// TIA Portal project "StdS71500PLCRack" (V17)

(* hardware
DEVICE "S7-1500/ET200MP-Station_1"  S7-1500 station
   slot 0: "Profilschiene_0"  Rack  6ES7 590-1***0-0AA0
   slot 1: "PLC_1"  CPU 1516-3 PN/DP  6ES7 516-3AN01-0AB0  V2.6
      slot 3: "CPU-Display_1"  6ES7591-1BA00-0AA0
      slot 32768: "PROFINET-Schnittstelle_1"  X1
      slot 33024: "PROFINET-Schnittstelle_2"  X2
      slot 33280: "DP-Schnittstelle_1"  X3
   slot 2: "DI 32x24VDC HF_1"  DI 32x24VDC HF  6ES7 521-1BL00-0AB0  V2.0
   slot 3: "DQ 32x24VDC/0.5A ST_1"  DQ 32x24VDC/0.5A ST  6ES7 522-1BL00-0AB0  V2.0
   slot 4: "AI 8xU/I/RTD/TC ST_1"  AI 8xU/I/RTD/TC ST  6ES7 531-7KF00-0AB0  V2.0
   slot 5: "AQ 4xU/I ST_1"  AQ 4xU/I ST  6ES7 532-5HD00-0AB0  V2.0
DEVICE "HMI_1"  TP700 Comfort
   slot 0: "HMI_1"  TP700 Comfort  6AV2 124-0GC01-0AX0  17.0.0.0
   slot 1: "HMI_RT_1"  TP700 Comfort  6AV2 124-0GC01-0AX0  17.0.0.0
   slot 5: "HMI_1.IE_CP_1"  PROFINET Interface  17.0.0.0
      slot 1: "PROFINET Interface_1"  PROFINET Interface
         slot 1: "Port_1"  Port
         slot 2: "Port_2"  Port
   slot 7: "HMI_1.MPI/DP_CP_1"  MPI/DP Interface  17.0.0.0
*)

// ===== PLC "PLC_1"  CPU 1516-3 PN/DP =====

VAR_GLOBAL   // PLC tag table "Standard-Variablentabelle"
   "System_Byte" AT %MB100 : Byte;
   "FirstScan" AT %M100.0 : Bool;
   "DiagStatusUpdate" AT %M100.1 : Bool;
   "AlwaysTRUE" AT %M100.2 : Bool;
   "AlwaysFALSE" AT %M100.3 : Bool;
   "Clock_Byte" AT %MB200 : Byte;
   "Clock_10Hz" AT %M200.0 : Bool;
   "Clock_5Hz" AT %M200.1 : Bool;
   "Clock_2.5Hz" AT %M200.2 : Bool;
   "Clock_2Hz" AT %M200.3 : Bool;
   "Clock_1.25Hz" AT %M200.4 : Bool;
   "Clock_1Hz" AT %M200.5 : Bool;
   "Clock_0.625Hz" AT %M200.6 : Bool;
   "Clock_0.5Hz" AT %M200.7 : Bool;
   "Tag_1" AT %M10.0 : Bool;
   "Tag_2" AT %M10.1 : Bool;
   "Tag_3" AT %M10.2 : Bool;
   "Tag_4" AT %M10.3 : Bool;
   "Tag_5" AT %M10.4 : Bool;
   "Tag_6" AT %M10.5 : Bool;
   "Tag_7" AT %M10.6 : Bool;
   "Tag_8" AT %M10.7 : Bool;
   "temp_AUTO_B" AT %M300.5 : Bool;
   "A_W_Testing" AT %M300.0 : Bool;
   "ACK_Status" AT %M300.2 : Bool;
   "Tag_11" AT %M300.3 : Bool;
   "Tag_9" AT %M300.7 : Bool;
   "Tag_10" AT %M11.0 : Bool;
   "Tag_12" AT %M11.1 : Bool;
   "Tag_13" AT %M11.2 : Bool;
END_VAR

DATA_BLOCK "PainMix_DB"   // DB1
{ S7_Optimized_Access := 'TRUE' }
VERSION : 0.1
   VAR
      Agitator_MainT : Int;
      Sol_1_Switch : Bool;
      Sol_1_Pipe1 : Int;
      Sol_1_Pipe2 : Int;
      RED_Pipe : Int;
      GREEN_Pipe : Int;
      BLUE_Pipe : Int;
      Control_Mode : Bool := false;
      Sol_1_ValveCont : Bool;
      Sol_1_Valve_Status : Bool;
      Sol_2_Valve_Status : Bool;
      Red_Valve_Status : Bool;
      Green_Valve_Status : Bool;
      Blue_Valve_Status : Bool;
      MainTank_Mixer_Status : Bool;
      Sol_2_ValveCont : Bool;
      Red_ValveCont : Bool;
      Green_ValveCont : Bool;
      Blue_ValveCont : Bool;
      Red_P_Rotor : Int;
      Green_P_Rotor : Int;
      Blue_P_Rotor : Int;
      Red_Tank_Level : Int := 40;
      Blue_Tank_Level : Int := 40;
      Green_Tank_Level : Int := 40;
      Sol_1_Tank_Level : Int := 40;
      Sol_2_Tank_Level : Int := 40;
      MainTank_Mixer_Cont : Bool;
      MainTank_Tank_Level : Int := 40;
      AUTO_Mode : Bool;
      AUTO_Mode_Prior : Int;
      temp_Auto_1 : Bool;
      Alarm_ACK : Bool;
   END_VAR
BEGIN
END_DATA_BLOCK

DATA_BLOCK "Paramters_Paint_Mix"   // DB7
{ S7_Optimized_Access := 'TRUE' }
VERSION : 0.1
   VAR
      ResinE_Flow_Act : Real := 1.6;
      ResinE_Flow_Set : Real := 1.8;
      Defoaming_Set : Real := 3.6;
      "Gloss Ratio_Set" : Real := 34.5;
      Binder_Flow_Act : Real := 2.2;
      Binder_Flow_Set : Real := 2.5;
      Level_Set_R : Real := 13.5;
      Level_Set_G : Real := 13.5;
      Level_Set_B : Real := 13.5;
      Flowrate_Set_R : Real := 3.1;
      Flowrate_Set_G : Real := 3.1;
      Flowrate_Set_B : Real := 3.1;
      Viscosity_Set_R : Real := 2.1;
      Viscosity_Set_G : Real := 2.7;
      Viscosity_Set_B : Real := 3.1;
      Density_Set_R : Real := 1.4;
      Density_Set_G : Real := 1.5;
      Density_Set_B : Real := 1.7;
      Temperature_Set_R : Real := 88.5;
      Temperature_Set_G : Real := 88.5;
      Temperature_Set_B : Real := 88.5;
      Pressure_Set_R : Real := 6.6;
      Pressure_Set_G : Real := 6.6;
      Pressure_Set_B : Real := 6.6;
      MixingSpeed_Set_MT : Real := 33.5;
      pH_MT : Real := 8.7;
      Viscosity_Set_MT : Real := 2.9;
      Level_Set_MT : Real := 17.0;
      Act_Red_Tank_Temp : Real := 73.5;
      Act_Green_Tank_Temp : Real := 76.2;
      Act_Blue_Tank_Temp : Real := 77.5;
      Act_Red_Tank_Press : Real := 5.3;
      Act_Green_Tank_Press : Real := 6.1;
      Act_Blue_Tank_Press : Real := 5.9;
      Recipe_Name : String := 'Pearl Gray';
      Recipe_ID : String := '001';
      Equip_ID : String := 'TN15112';
      Batch_ID : String := '052B';
      Batch_Size : String := '85 litr';
      Start_Time : String := '28/01/2025, 14:56:32';
      Alarm_1 : Bool;
      Alarm_2 : Bool;
      Warning_1 : Bool;
      Warning_2 : Bool;
      Warning_3 : Bool;
      "Common_A-W" : Bool;
      Language : Bool := false;
      Button_Language : Bool;
      MainOverview : Bool;
      Parameters : Bool;
      RecipeM : Bool;
      UserM : Bool;
      AlarmSt : Bool;
      IOSt : Bool;
   END_VAR
BEGIN
END_DATA_BLOCK

DATA_BLOCK "DI"   // DB8
{ S7_Optimized_Access := 'TRUE' }
VERSION : 0.1
   VAR
      "I0.0" : Bool;
      "I0.1" : Bool := true;
      "I0.2" : Bool;
      "I0.3" : Bool := true;
      "I0.4" : Bool;
      "I0.5" : Bool;
      "I0.6" : Bool := true;
      "I0.7" : Bool;
      "I1.0" : Bool;
      "I1.1" : Bool;
      "I1.2" : Bool;
      "I1.3" : Bool := true;
      "I1.4" : Bool;
      "I1.5" : Bool;
      "I1.6" : Bool;
      "I1.7" : Bool := true;
      "I2.0" : Bool := true;
      "I2.1" : Bool;
      "I2.2" : Bool;
      "I2.3" : Bool := true;
   END_VAR
BEGIN
END_DATA_BLOCK

DATA_BLOCK "DO"   // DB9
{ S7_Optimized_Access := 'TRUE' }
VERSION : 0.1
   VAR
      "Q0.0" : Bool;
      "Q0.1" : Bool;
      "Q0.2" : Bool;
      "Q0.3" : Bool;
      "Q0.4" : Bool;
      "Q0.5" : Bool;
      "Q0.6" : Bool;
      "Q0.7" : Bool;
      "Q1.0" : Bool;
      "Q1.1" : Bool;
      "Q1.2" : Bool;
      "Q1.3" : Bool;
      "Q1.4" : Bool;
      "Q1.5" : Bool;
      "Q1.6" : Bool;
      "Q1.7" : Bool := true;
      "Q2.0" : Bool;
      "Q2.1" : Bool;
      "Q2.2" : Bool := true;
      "Q2.3" : Bool := true;
   END_VAR
BEGIN
END_DATA_BLOCK

DATA_BLOCK "Recipe"   // DB10
{ S7_Optimized_Access := 'TRUE' }
VERSION : 0.1
   VAR
      "Pigment Concentration" : Real;
      "Resin Type and Ratio" : Real;
      "Solvent Composition" : Real;
      "Additive Ratios" : Real;
      "Drying Agent Ratio" : Real;
      "Viscosity Target" : Real;
      "Gloss Level" : Real;
      "pH Control Range" : Real;
      "Mixing Time" : Real;
      "Curing Agent Proportion" : Real;
      Recipe_Name : String;
   END_VAR
BEGIN
END_DATA_BLOCK

// folder: System blocks/Program resources

DATA_BLOCK "IEC_Timer_0_DB"   // DB2
{ S7_Optimized_Access := 'TRUE' }
AUTHOR : Simatic
FAMILY : IEC
NAME : IEC_TMR
VERSION : 1.0
// stored: InstanceOfName IEC_TIMER
"IEC_TIMER"
BEGIN
END_DATA_BLOCK

DATA_BLOCK "IEC_Timer_0_DB_1"   // DB3
{ S7_Optimized_Access := 'TRUE' }
AUTHOR : Simatic
FAMILY : IEC
NAME : IEC_TMR
VERSION : 1.0
// stored: InstanceOfName IEC_TIMER
"IEC_TIMER"
BEGIN
END_DATA_BLOCK

DATA_BLOCK "IEC_Timer_0_DB_2"   // DB4
{ S7_Optimized_Access := 'TRUE' }
AUTHOR : Simatic
FAMILY : IEC
NAME : IEC_TMR
VERSION : 1.0
// stored: InstanceOfName IEC_TIMER
"IEC_TIMER"
BEGIN
END_DATA_BLOCK

DATA_BLOCK "IEC_Timer_0_DB_3"   // DB5
{ S7_Optimized_Access := 'TRUE' }
AUTHOR : Simatic
FAMILY : IEC
NAME : IEC_TMR
VERSION : 1.0
// stored: InstanceOfName IEC_TIMER
"IEC_TIMER"
BEGIN
END_DATA_BLOCK

DATA_BLOCK "IEC_Timer_0_DB_4"   // DB6
{ S7_Optimized_Access := 'TRUE' }
AUTHOR : Simatic
FAMILY : IEC
NAME : IEC_TMR
VERSION : 1.0
// stored: InstanceOfName IEC_TIMER
"IEC_TIMER"
BEGIN
END_DATA_BLOCK

DATA_BLOCK "IEC_Timer_0_DB_5"   // DB11
{ S7_Optimized_Access := 'TRUE' }
AUTHOR : Simatic
FAMILY : IEC
NAME : IEC_TMR
VERSION : 1.0
// stored: InstanceOfName IEC_TIMER
"IEC_TIMER"
BEGIN
END_DATA_BLOCK

DATA_BLOCK "IEC_Counter_0_DB"   // DB12
{ S7_Optimized_Access := 'TRUE' }
AUTHOR : Simatic
FAMILY : IEC
NAME : CNTR
VERSION : 1.0
// stored: InstanceOfName IEC_COUNTER
"IEC_COUNTER"
BEGIN
END_DATA_BLOCK

DATA_BLOCK "IEC_Timer_0_DB_6"   // DB13
{ S7_Optimized_Access := 'TRUE' }
AUTHOR : Simatic
FAMILY : IEC
NAME : IEC_TMR
VERSION : 1.0
// stored: InstanceOfName IEC_TIMER
"IEC_TIMER"
BEGIN
END_DATA_BLOCK

// folder: (top level)

ORGANIZATION_BLOCK "Main"   // OB1, LAD, ProgramCycle
TITLE = "Main Program Sweep (Cycle)"
{ S7_Optimized_Access := 'TRUE' }
VERSION : 0.1
   VAR_INPUT
      Initial_Call : Bool;   // Initial call of this OB
      Remanence : Bool;   // =True, if remanent data are available
   END_VAR
   VAR_TEMP   // added for the SCL form of the ladder/FBD networks
      _w1 : Bool;
      _w2 : Bool;
   END_VAR
BEGIN

REGION Network 1: AUTO Sequence Logic
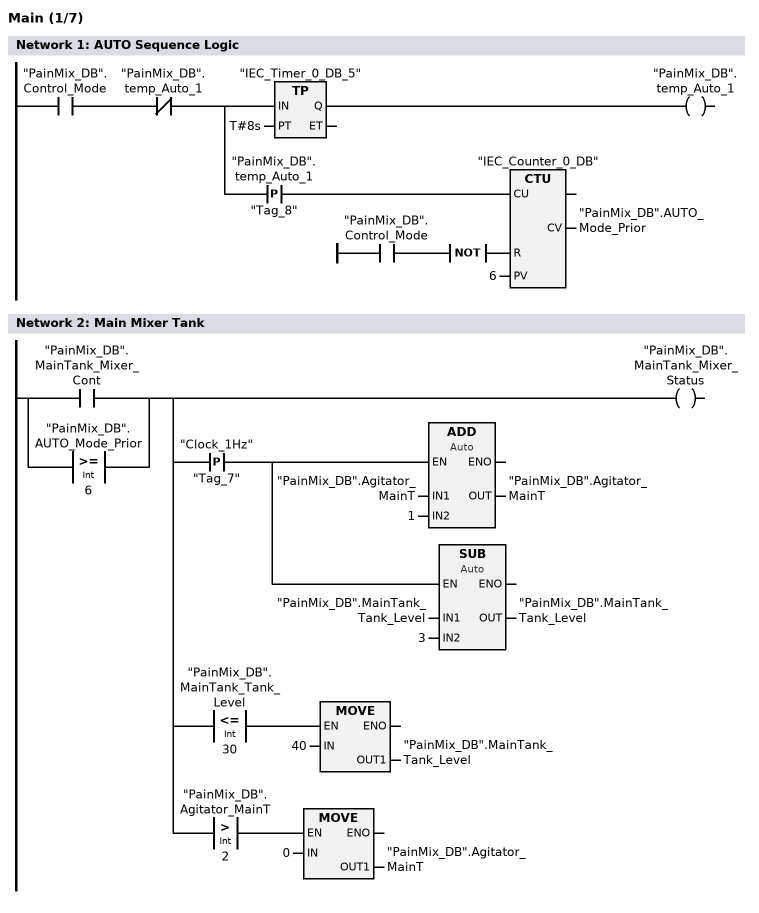
   #_w1 := "PainMix_DB".Control_Mode AND NOT "PainMix_DB".temp_Auto_1;
   "IEC_Timer_0_DB_5".TP(IN := #_w1, PT := T#8s);
   "PainMix_DB".temp_Auto_1 := "IEC_Timer_0_DB_5".Q;
   #_w2 := #_w1 AND "PainMix_DB".temp_Auto_1 AND NOT "Tag_8";   // rising edge of "PainMix_DB".temp_Auto_1
   "Tag_8" := "PainMix_DB".temp_Auto_1;
   "IEC_Counter_0_DB".CTU(CU := #_w2,
                          R := NOT "PainMix_DB".Control_Mode,
                          PV := 6,
                          CV => "PainMix_DB".AUTO_Mode_Prior);
END_REGION

REGION Network 2: Main Mixer Tank
   RUNG wire#powerrail
      Contact( "PainMix_DB".MainTank_Mixer_Cont )
      wire#w1
      Coil( "PainMix_DB".MainTank_Mixer_Status )
   END_RUNG
   RUNG wire#powerrail
      { S7_Templates := "SrcType := Int" } GE_Contact(in1 := "PainMix_DB".AUTO_Mode_Prior, in2 := 6)
   END_RUNG wire#w1
   RUNG wire#w1
      P_Contact(operand := "Clock_1Hz", bit := "Tag_7")
      wire#w2
      Add(in1 := "PainMix_DB".Agitator_MainT, in2 := 1, out => "PainMix_DB".Agitator_MainT)
   END_RUNG
   RUNG wire#w2
      Sub(in1 := "PainMix_DB".MainTank_Tank_Level, in2 := 3, out => "PainMix_DB".MainTank_Tank_Level)
   END_RUNG
   RUNG wire#w1
      { S7_Templates := "SrcType := Int" } LE_Contact(in1 := "PainMix_DB".MainTank_Tank_Level, in2 := 30)
      Move(in := 40, out1 => "PainMix_DB".MainTank_Tank_Level)
   END_RUNG
   RUNG wire#w1
      { S7_Templates := "SrcType := Int" } GT_Contact(in1 := "PainMix_DB".Agitator_MainT, in2 := 2)
      Move(in := 0, out1 => "PainMix_DB".Agitator_MainT)
   END_RUNG
   // the same network as SCL:
   "PainMix_DB".MainTank_Mixer_Status := "PainMix_DB".MainTank_Mixer_Cont OR ("PainMix_DB".AUTO_Mode_Prior >= 6);
   #_w1 := "PainMix_DB".MainTank_Mixer_Status AND "Clock_1Hz" AND NOT "Tag_7";   // rising edge of "Clock_1Hz"
   "Tag_7" := "Clock_1Hz";
   IF #_w1 THEN
       "PainMix_DB".Agitator_MainT := "PainMix_DB".Agitator_MainT + 1;
       "PainMix_DB".MainTank_Tank_Level := "PainMix_DB".MainTank_Tank_Level - 3;
   END_IF;
   IF "PainMix_DB".MainTank_Mixer_Status AND ("PainMix_DB".MainTank_Tank_Level <= 30) THEN
       "PainMix_DB".MainTank_Tank_Level := 40;
   END_IF;
   IF "PainMix_DB".MainTank_Mixer_Status AND ("PainMix_DB".Agitator_MainT > 2) THEN
       "PainMix_DB".Agitator_MainT := 0;
   END_IF;
END_REGION

REGION Network 3: Resin Solution
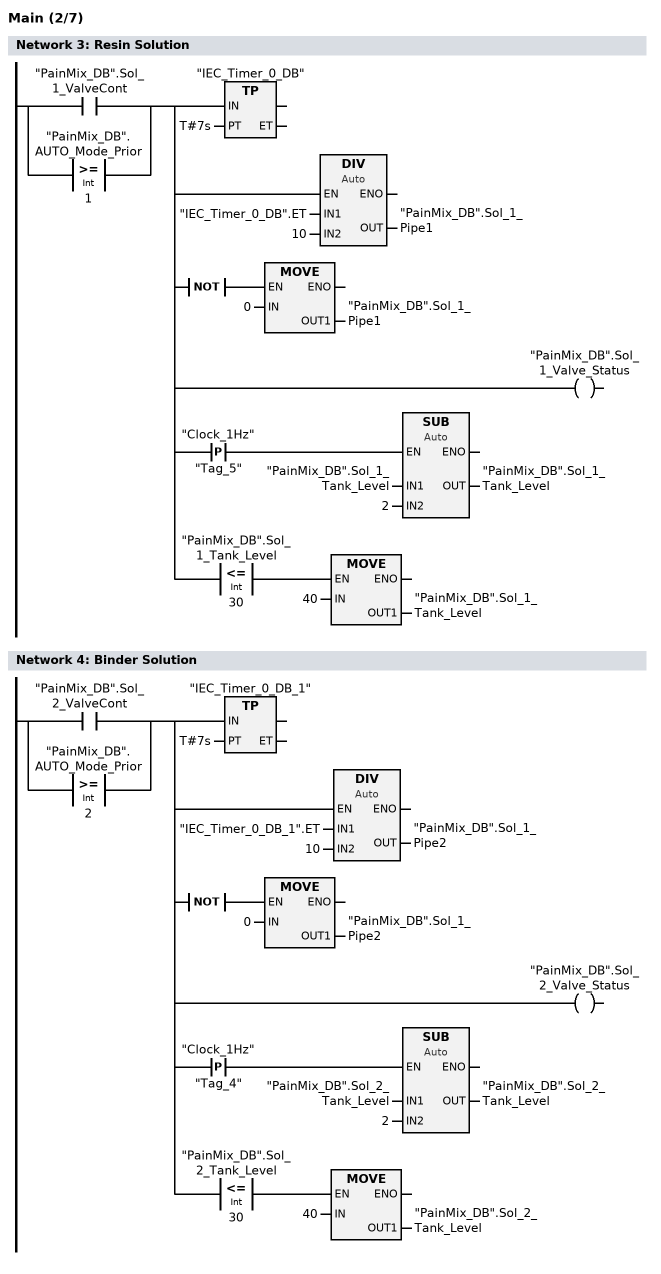
   #_w1 := "PainMix_DB".Sol_1_ValveCont OR ("PainMix_DB".AUTO_Mode_Prior >= 1);
   "IEC_Timer_0_DB".TP(IN := #_w1, PT := T#7s);
   IF #_w1 THEN "PainMix_DB".Sol_1_Pipe1 := "IEC_Timer_0_DB".ET / 10; END_IF;
   IF NOT #_w1 THEN "PainMix_DB".Sol_1_Pipe1 := 0; END_IF;
   "PainMix_DB".Sol_1_Valve_Status := #_w1;
   #_w2 := #_w1 AND "Clock_1Hz" AND NOT "Tag_5";   // rising edge of "Clock_1Hz"
   "Tag_5" := "Clock_1Hz";
   IF #_w2 THEN "PainMix_DB".Sol_1_Tank_Level := "PainMix_DB".Sol_1_Tank_Level - 2; END_IF;
   IF #_w1 AND ("PainMix_DB".Sol_1_Tank_Level <= 30) THEN "PainMix_DB".Sol_1_Tank_Level := 40; END_IF;
END_REGION

REGION Network 4: Binder Solution
   #_w1 := "PainMix_DB".Sol_2_ValveCont OR ("PainMix_DB".AUTO_Mode_Prior >= 2);
   "IEC_Timer_0_DB_1".TP(IN := #_w1, PT := T#7s);
   IF #_w1 THEN "PainMix_DB".Sol_1_Pipe2 := "IEC_Timer_0_DB_1".ET / 10; END_IF;
   IF NOT #_w1 THEN "PainMix_DB".Sol_1_Pipe2 := 0; END_IF;
   "PainMix_DB".Sol_2_Valve_Status := #_w1;
   #_w2 := #_w1 AND "Clock_1Hz" AND NOT "Tag_4";   // rising edge of "Clock_1Hz"
   "Tag_4" := "Clock_1Hz";
   IF #_w2 THEN "PainMix_DB".Sol_2_Tank_Level := "PainMix_DB".Sol_2_Tank_Level - 2; END_IF;
   IF #_w1 AND ("PainMix_DB".Sol_2_Tank_Level <= 30) THEN "PainMix_DB".Sol_2_Tank_Level := 40; END_IF;
END_REGION

REGION Network 5: RED
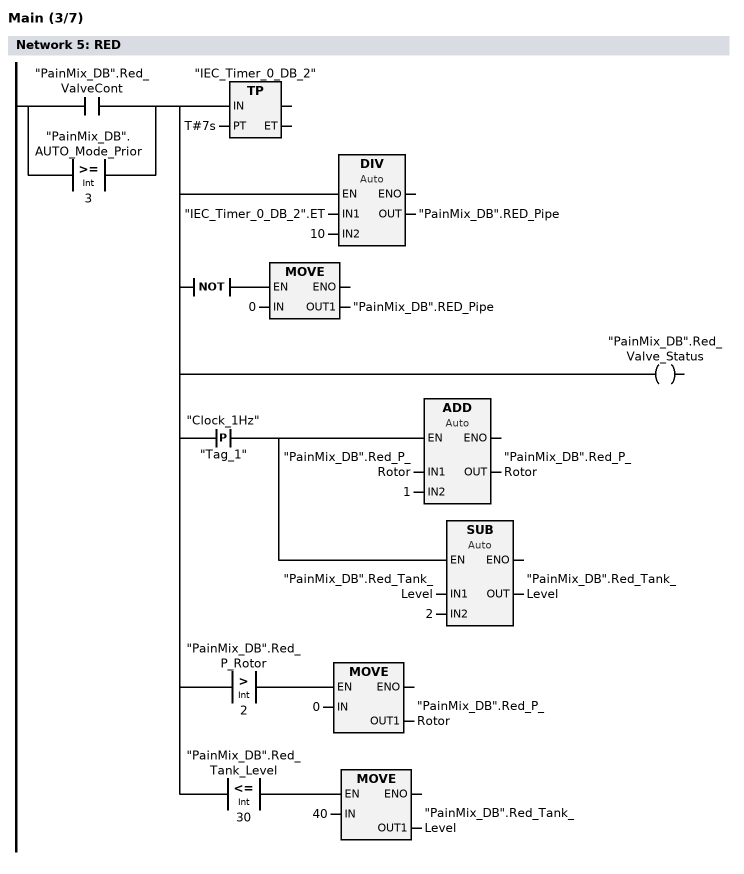
   #_w1 := "PainMix_DB".Red_ValveCont OR ("PainMix_DB".AUTO_Mode_Prior >= 3);
   "IEC_Timer_0_DB_2".TP(IN := #_w1, PT := T#7s);
   IF #_w1 THEN "PainMix_DB".RED_Pipe := "IEC_Timer_0_DB_2".ET / 10; END_IF;
   IF NOT #_w1 THEN "PainMix_DB".RED_Pipe := 0; END_IF;
   "PainMix_DB".Red_Valve_Status := #_w1;
   #_w2 := #_w1 AND "Clock_1Hz" AND NOT "Tag_1";   // rising edge of "Clock_1Hz"
   "Tag_1" := "Clock_1Hz";
   IF #_w2 THEN
       "PainMix_DB".Red_P_Rotor := "PainMix_DB".Red_P_Rotor + 1;
       "PainMix_DB".Red_Tank_Level := "PainMix_DB".Red_Tank_Level - 2;
   END_IF;
   IF #_w1 AND ("PainMix_DB".Red_P_Rotor > 2) THEN "PainMix_DB".Red_P_Rotor := 0; END_IF;
   IF #_w1 AND ("PainMix_DB".Red_Tank_Level <= 30) THEN "PainMix_DB".Red_Tank_Level := 40; END_IF;
END_REGION

REGION Network 6: GREEN
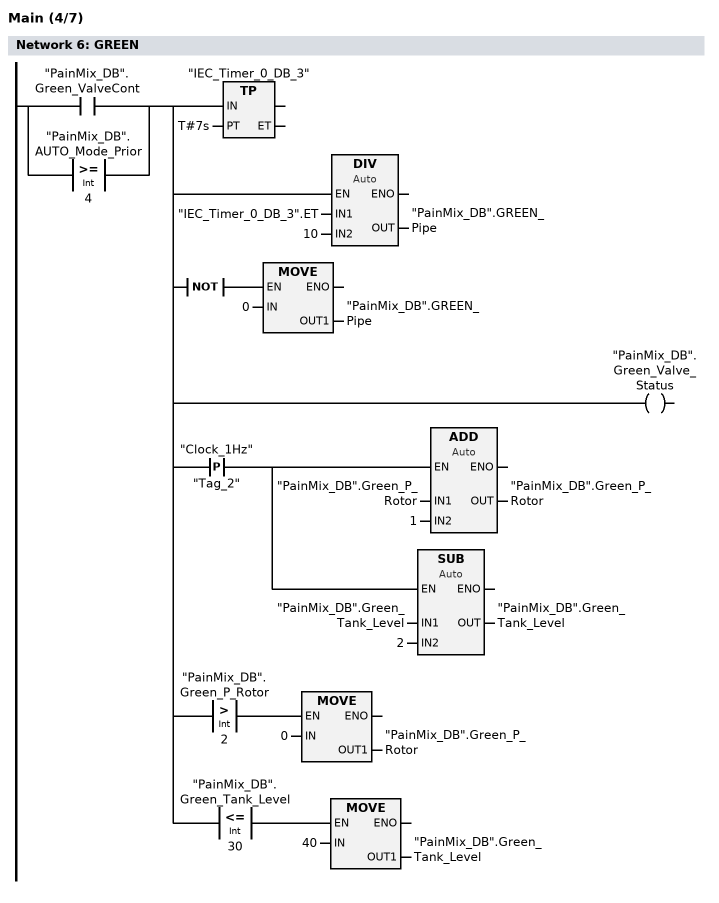
   #_w1 := "PainMix_DB".Green_ValveCont OR ("PainMix_DB".AUTO_Mode_Prior >= 4);
   "IEC_Timer_0_DB_3".TP(IN := #_w1, PT := T#7s);
   IF #_w1 THEN "PainMix_DB".GREEN_Pipe := "IEC_Timer_0_DB_3".ET / 10; END_IF;
   IF NOT #_w1 THEN "PainMix_DB".GREEN_Pipe := 0; END_IF;
   "PainMix_DB".Green_Valve_Status := #_w1;
   #_w2 := #_w1 AND "Clock_1Hz" AND NOT "Tag_2";   // rising edge of "Clock_1Hz"
   "Tag_2" := "Clock_1Hz";
   IF #_w2 THEN
       "PainMix_DB".Green_P_Rotor := "PainMix_DB".Green_P_Rotor + 1;
       "PainMix_DB".Green_Tank_Level := "PainMix_DB".Green_Tank_Level - 2;
   END_IF;
   IF #_w1 AND ("PainMix_DB".Green_P_Rotor > 2) THEN "PainMix_DB".Green_P_Rotor := 0; END_IF;
   IF #_w1 AND ("PainMix_DB".Green_Tank_Level <= 30) THEN "PainMix_DB".Green_Tank_Level := 40; END_IF;
END_REGION

REGION Network 7: BLUE
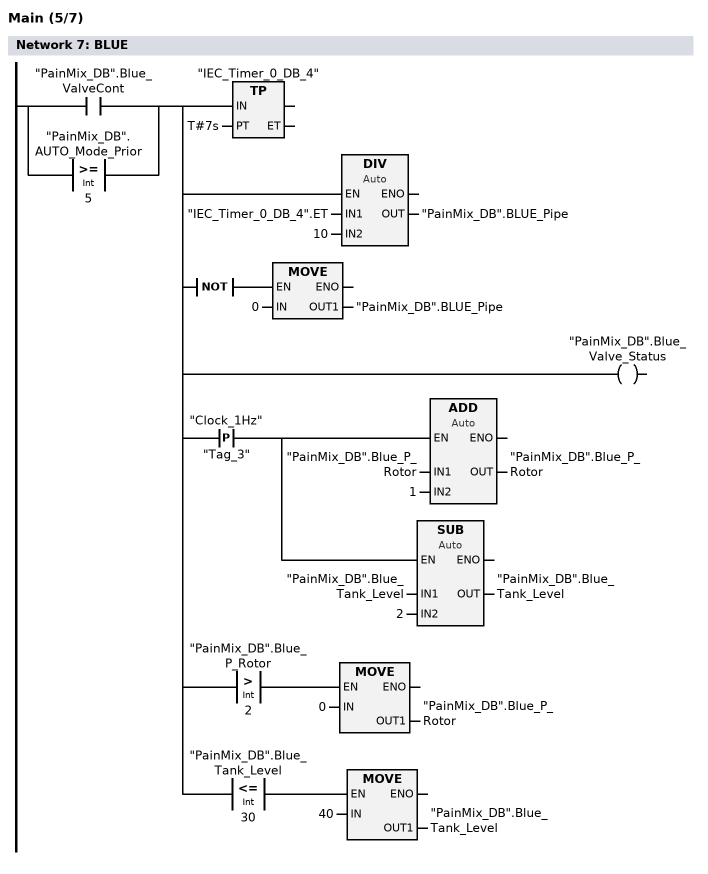
   #_w1 := "PainMix_DB".Blue_ValveCont OR ("PainMix_DB".AUTO_Mode_Prior >= 5);
   "IEC_Timer_0_DB_4".TP(IN := #_w1, PT := T#7s);
   IF #_w1 THEN "PainMix_DB".BLUE_Pipe := "IEC_Timer_0_DB_4".ET / 10; END_IF;
   IF NOT #_w1 THEN "PainMix_DB".BLUE_Pipe := 0; END_IF;
   "PainMix_DB".Blue_Valve_Status := #_w1;
   #_w2 := #_w1 AND "Clock_1Hz" AND NOT "Tag_3";   // rising edge of "Clock_1Hz"
   "Tag_3" := "Clock_1Hz";
   IF #_w2 THEN
       "PainMix_DB".Blue_P_Rotor := "PainMix_DB".Blue_P_Rotor + 1;
       "PainMix_DB".Blue_Tank_Level := "PainMix_DB".Blue_Tank_Level - 2;
   END_IF;
   IF #_w1 AND ("PainMix_DB".Blue_P_Rotor > 2) THEN "PainMix_DB".Blue_P_Rotor := 0; END_IF;
   IF #_w1 AND ("PainMix_DB".Blue_Tank_Level <= 30) THEN "PainMix_DB".Blue_Tank_Level := 40; END_IF;
END_REGION

REGION Network 8: Flucuation of Temp & Press of Tanks
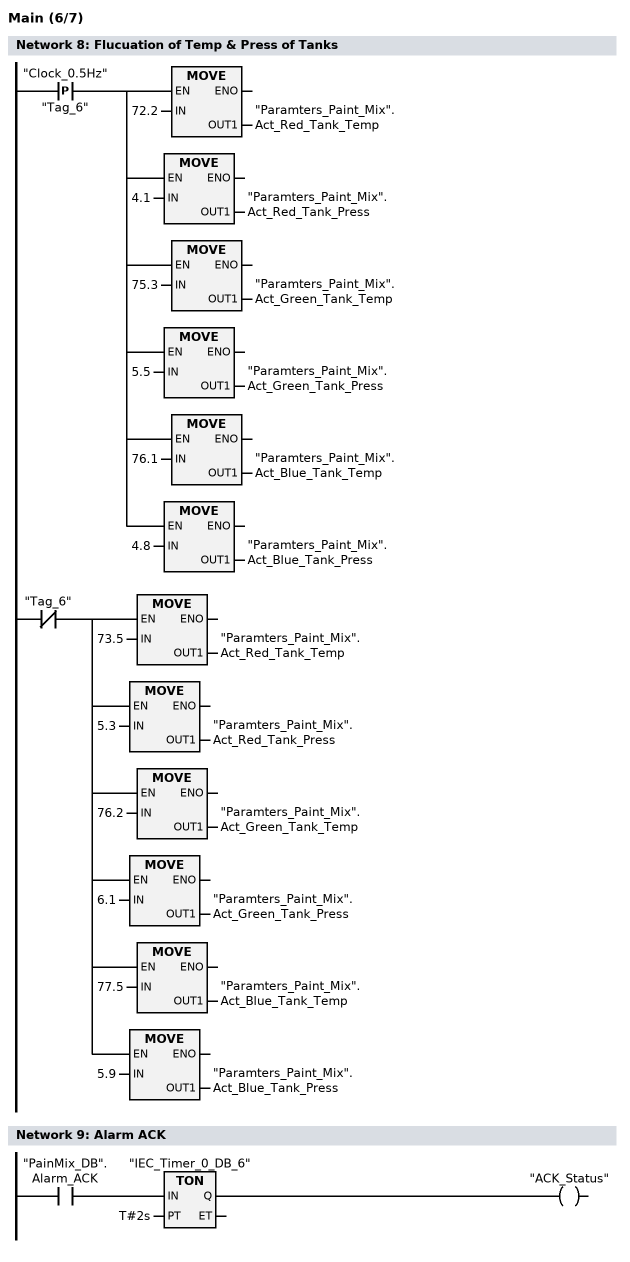
   RUNG wire#powerrail
      P_Contact(operand := "Clock_0.5Hz", bit := "Tag_6")
      wire#w1
      Move(in := 72.2, out1 => "Paramters_Paint_Mix".Act_Red_Tank_Temp)
   END_RUNG
   RUNG wire#w1
      Move(in := 4.1, out1 => "Paramters_Paint_Mix".Act_Red_Tank_Press)
   END_RUNG
   RUNG wire#w1
      Move(in := 75.3, out1 => "Paramters_Paint_Mix".Act_Green_Tank_Temp)
   END_RUNG
   RUNG wire#w1
      Move(in := 5.5, out1 => "Paramters_Paint_Mix".Act_Green_Tank_Press)
   END_RUNG
   RUNG wire#w1
      Move(in := 76.1, out1 => "Paramters_Paint_Mix".Act_Blue_Tank_Temp)
   END_RUNG
   RUNG wire#w1
      Move(in := 4.8, out1 => "Paramters_Paint_Mix".Act_Blue_Tank_Press)
   END_RUNG
   RUNG wire#powerrail
      I_Contact( "Tag_6" )
      wire#w2
      Move(in := 73.5, out1 => "Paramters_Paint_Mix".Act_Red_Tank_Temp)
   END_RUNG
   RUNG wire#w2
      Move(in := 5.3, out1 => "Paramters_Paint_Mix".Act_Red_Tank_Press)
   END_RUNG
   RUNG wire#w2
      Move(in := 76.2, out1 => "Paramters_Paint_Mix".Act_Green_Tank_Temp)
   END_RUNG
   RUNG wire#w2
      Move(in := 6.1, out1 => "Paramters_Paint_Mix".Act_Green_Tank_Press)
   END_RUNG
   RUNG wire#w2
      Move(in := 77.5, out1 => "Paramters_Paint_Mix".Act_Blue_Tank_Temp)
   END_RUNG
   RUNG wire#w2
      Move(in := 5.9, out1 => "Paramters_Paint_Mix".Act_Blue_Tank_Press)
   END_RUNG
   // the same network as SCL:
   #_w1 := "Clock_0.5Hz" AND NOT "Tag_6";   // rising edge of "Clock_0.5Hz"
   "Tag_6" := "Clock_0.5Hz";
   IF #_w1 THEN
       "Paramters_Paint_Mix".Act_Red_Tank_Temp := 72.2;
       "Paramters_Paint_Mix".Act_Red_Tank_Press := 4.1;
       "Paramters_Paint_Mix".Act_Green_Tank_Temp := 75.3;
       "Paramters_Paint_Mix".Act_Green_Tank_Press := 5.5;
       "Paramters_Paint_Mix".Act_Blue_Tank_Temp := 76.1;
       "Paramters_Paint_Mix".Act_Blue_Tank_Press := 4.8;
   END_IF;
   IF NOT "Tag_6" THEN
       "Paramters_Paint_Mix".Act_Red_Tank_Temp := 73.5;
       "Paramters_Paint_Mix".Act_Red_Tank_Press := 5.3;
       "Paramters_Paint_Mix".Act_Green_Tank_Temp := 76.2;
       "Paramters_Paint_Mix".Act_Green_Tank_Press := 6.1;
       "Paramters_Paint_Mix".Act_Blue_Tank_Temp := 77.5;
       "Paramters_Paint_Mix".Act_Blue_Tank_Press := 5.9;
   END_IF;
END_REGION

REGION Network 9: Alarm ACK
   "IEC_Timer_0_DB_6".TON(IN := "PainMix_DB".Alarm_ACK, PT := T#2s);
   "ACK_Status" := "IEC_Timer_0_DB_6".Q;
END_REGION

REGION Network 10: Alarm - Warning --- ON
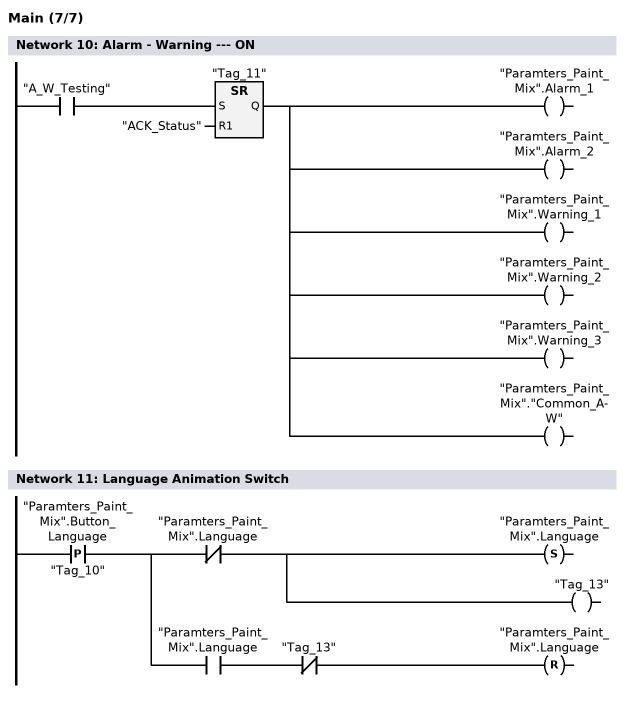
   RUNG wire#powerrail
      Contact( "A_W_Testing" )
      S_SR(operand := "Tag_11", r1 := "ACK_Status")
      wire#w1
      Coil( "Paramters_Paint_Mix".Alarm_1 )
   END_RUNG
   RUNG wire#w1
      Coil( "Paramters_Paint_Mix".Alarm_2 )
   END_RUNG
   RUNG wire#w1
      Coil( "Paramters_Paint_Mix".Warning_1 )
   END_RUNG
   RUNG wire#w1
      Coil( "Paramters_Paint_Mix".Warning_2 )
   END_RUNG
   RUNG wire#w1
      Coil( "Paramters_Paint_Mix".Warning_3 )
   END_RUNG
   RUNG wire#w1
      Coil( "Paramters_Paint_Mix"."Common_A-W" )
   END_RUNG
   // the same network as SCL:
   IF "A_W_Testing" THEN
       "Tag_11" := TRUE;   // SR flip-flop
   END_IF;
   IF "ACK_Status" THEN "Tag_11" := FALSE; END_IF;
   "Paramters_Paint_Mix".Alarm_1 := "Tag_11";
   "Paramters_Paint_Mix".Alarm_2 := "Tag_11";
   "Paramters_Paint_Mix".Warning_1 := "Tag_11";
   "Paramters_Paint_Mix".Warning_2 := "Tag_11";
   "Paramters_Paint_Mix".Warning_3 := "Tag_11";
   "Paramters_Paint_Mix"."Common_A-W" := "Tag_11";
END_REGION

REGION Network 11: Language Animation Switch
   RUNG wire#powerrail
      P_Contact(operand := "Paramters_Paint_Mix".Button_Language, bit := "Tag_10")
      wire#w1
      I_Contact( "Paramters_Paint_Mix".Language )
      wire#w2
      S_Coil( "Paramters_Paint_Mix".Language )
   END_RUNG
   RUNG wire#w2
      Coil( "Tag_13" )
   END_RUNG
   RUNG wire#w1
      Contact( "Paramters_Paint_Mix".Language )
      I_Contact( "Tag_13" )
      R_Coil( "Paramters_Paint_Mix".Language )
   END_RUNG
   // the same network as SCL:
   #_w1 := "Paramters_Paint_Mix".Button_Language AND NOT "Tag_10";   // rising edge of "Paramters_Paint_Mix".Button_Language
   "Tag_10" := "Paramters_Paint_Mix".Button_Language;
   #_w2 := #_w1 AND NOT "Paramters_Paint_Mix".Language;
   IF #_w2 THEN "Paramters_Paint_Mix".Language := TRUE; END_IF;
   "Tag_13" := #_w2;
   IF #_w1 AND "Paramters_Paint_Mix".Language AND NOT "Tag_13" THEN
       "Paramters_Paint_Mix".Language := FALSE;
   END_IF;
END_REGION
END_ORGANIZATION_BLOCK

(* ===== HMI "HMI_RT_1" =====
system functions are stored by id; their names below are inferred from use
connection "HMI_Connection_1": ETHERNET, S7_1500_OMS

HMI tags "Default tag table"
   "PainMix_DB_Sol_1_Switch" : Bool = PLC PainMix_DB.Sol_1_Switch, 1 s
   "PainMix_DB_Sol_1_Pipe1" : Int = PLC PainMix_DB.Sol_1_Pipe1, 1 s
   "PainMix_DB_Sol_1_Pipe2" : Int = PLC PainMix_DB.Sol_1_Pipe2, 1 s
   "PainMix_DB_RED_Pipe" : Int = PLC PainMix_DB.RED_Pipe, 1 s
   "PainMix_DB_GREEN_Pipe" : Int = PLC PainMix_DB.GREEN_Pipe, 1 s
   "PainMix_DB_BLUE_Pipe" : Int = PLC PainMix_DB.BLUE_Pipe, 1 s
   "PainMix_DB_Control_Mode" : Bool = PLC PainMix_DB.Control_Mode, 1 s
   "PainMix_DB_Sol_1_ValveCont" : Bool = PLC PainMix_DB.Sol_1_ValveCont, 1 s
   "PainMix_DB_Sol_1_Valve_Status" : Bool = PLC PainMix_DB.Sol_1_Valve_Status, 1 s
   "PainMix_DB_Sol_2_Valve_Status" : Bool = PLC PainMix_DB.Sol_2_Valve_Status, 1 s
   "PainMix_DB_Red_Valve_Status" : Bool = PLC PainMix_DB.Red_Valve_Status, 1 s
   "PainMix_DB_Green_Valve_Status" : Bool = PLC PainMix_DB.Green_Valve_Status, 1 s
   "PainMix_DB_Blue_Valve_Status" : Bool = PLC PainMix_DB.Blue_Valve_Status, 1 s
   "PainMix_DB_MainTank_Mixer_Status" : Bool = PLC PainMix_DB.MainTank_Mixer_Status, 1 s
   "PainMix_DB_Sol_2_ValveCont" : Bool = PLC PainMix_DB.Sol_2_ValveCont, 1 s
   "PainMix_DB_Red_ValveCont" : Bool = PLC PainMix_DB.Red_ValveCont, 1 s
   "PainMix_DB_Green_ValveCont" : Bool = PLC PainMix_DB.Green_ValveCont, 1 s
   "PainMix_DB_Blue_ValveCont" : Bool = PLC PainMix_DB.Blue_ValveCont, 1 s
   "Paramters_Paint_Mix_ResinE_Flow_Act" : Real = PLC Paramters_Paint_Mix.ResinE_Flow_Act, 1 s
   "Paramters_Paint_Mix_ResinE_Flow_Set" : Real = PLC Paramters_Paint_Mix.ResinE_Flow_Set, 1 s
   "Paramters_Paint_Mix_Binder_Flow_Act" : Real = PLC Paramters_Paint_Mix.Binder_Flow_Act, 1 s
   "Paramters_Paint_Mix_Binder_Flow_Set" : Real = PLC Paramters_Paint_Mix.Binder_Flow_Set, 1 s
   "Paramters_Paint_Mix_Defoaming_Set" : Real = PLC Paramters_Paint_Mix.Defoaming_Set, 1 s
   "Paramters_Paint_Mix_Gloss Ratio_Set" : Real = PLC Paramters_Paint_Mix."Gloss Ratio_Set", 1 s
   "Paramters_Paint_Mix_Level_Set_R" : Real = PLC Paramters_Paint_Mix.Level_Set_R, 1 s
   "Paramters_Paint_Mix_Flowrate_Set_R" : Real = PLC Paramters_Paint_Mix.Flowrate_Set_R, 1 s
   "Paramters_Paint_Mix_Viscosity_Set_R" : Real = PLC Paramters_Paint_Mix.Viscosity_Set_R, 1 s
   "Paramters_Paint_Mix_Density_Set_R" : Real = PLC Paramters_Paint_Mix.Density_Set_R, 1 s
   "Paramters_Paint_Mix_Temperature_Set_R" : Real = PLC Paramters_Paint_Mix.Temperature_Set_R, 1 s
   "Paramters_Paint_Mix_Pressure_Set_R" : Real = PLC Paramters_Paint_Mix.Pressure_Set_R, 1 s
   "Paramters_Paint_Mix_MixingSpeed_Set_MT" : Real = PLC Paramters_Paint_Mix.MixingSpeed_Set_MT, 1 s
   "Paramters_Paint_Mix_pH_MT" : Real = PLC Paramters_Paint_Mix.pH_MT, 1 s
   "Paramters_Paint_Mix_Viscosity_Set_MT" : Real = PLC Paramters_Paint_Mix.Viscosity_Set_MT, 1 s
   "Paramters_Paint_Mix_Level_Set_MT" : Real = PLC Paramters_Paint_Mix.Level_Set_MT, 1 s
   "PainMix_DB_Red_P_Rotor" : Int = PLC PainMix_DB.Red_P_Rotor, 1 s
   "PainMix_DB_Green_P_Rotor" : Int = PLC PainMix_DB.Green_P_Rotor, 1 s
   "PainMix_DB_Blue_P_Rotor" : Int = PLC PainMix_DB.Blue_P_Rotor, 1 s
   "PainMix_DB_Red_Tank_Level" : Int = PLC PainMix_DB.Red_Tank_Level, 1 s
   "DI_I0.1" : Bool = PLC DI."I0.1", 1 s
   "DI_I0.2" : Bool = PLC DI."I0.2", 1 s
   "DI_I0.0" : Bool = PLC DI."I0.0", 1 s
   "DI_I0.4" : Bool = PLC DI."I0.4", 1 s
   "DI_I0.5" : Bool = PLC DI."I0.5", 1 s
   "DI_I0.6" : Bool = PLC DI."I0.6", 1 s
   "DI_I0.7" : Bool = PLC DI."I0.7", 1 s
   "DI_I1.0" : Bool = PLC DI."I1.0", 1 s
   "DI_I1.1" : Bool = PLC DI."I1.1", 1 s
   "DI_I1.2" : Bool = PLC DI."I1.2", 1 s
   "DI_I1.3" : Bool = PLC DI."I1.3", 1 s
   "DI_I1.4" : Bool = PLC DI."I1.4", 1 s
   "DI_I1.5" : Bool = PLC DI."I1.5", 1 s
   "DI_I1.6" : Bool = PLC DI."I1.6", 1 s
   "DI_I1.7" : Bool = PLC DI."I1.7", 1 s
   "DI_I2.0" : Bool = PLC DI."I2.0", 1 s
   "DI_I2.1" : Bool = PLC DI."I2.1", 1 s
   "DI_I2.2" : Bool = PLC DI."I2.2", 1 s
   "DI_I2.3" : Bool = PLC DI."I2.3", 1 s
   "DO_Q0.0" : Bool = PLC DO."Q0.0", 1 s
   "DO_Q0.1" : Bool = PLC DO."Q0.1", 1 s
   "DO_Q0.2" : Bool = PLC DO."Q0.2", 1 s
   "DO_Q0.3" : Bool = PLC DO."Q0.3", 1 s
   "DO_Q0.4" : Bool = PLC DO."Q0.4", 1 s
   "DO_Q0.5" : Bool = PLC DO."Q0.5", 1 s
   "DO_Q0.6" : Bool = PLC DO."Q0.6", 1 s
   "DO_Q0.7" : Bool = PLC DO."Q0.7", 1 s
   "DO_Q1.0" : Bool = PLC DO."Q1.0", 1 s
   "DO_Q1.1" : Bool = PLC DO."Q1.1", 1 s
   "DO_Q1.2" : Bool = PLC DO."Q1.2", 1 s
   "DO_Q1.3" : Bool = PLC DO."Q1.3", 1 s
   "DO_Q1.4" : Bool = PLC DO."Q1.4", 1 s
   "DO_Q1.5" : Bool = PLC DO."Q1.5", 1 s
   "DO_Q1.6" : Bool = PLC DO."Q1.6", 1 s
   "DO_Q1.7" : Bool = PLC DO."Q1.7", 1 s
   "DO_Q2.0" : Bool = PLC DO."Q2.0", 1 s
   "DO_Q2.1" : Bool = PLC DO."Q2.1", 1 s
   "DO_Q2.2" : Bool = PLC DO."Q2.2", 1 s
   "DO_Q2.3" : Bool = PLC DO."Q2.3", 1 s
   "Paramters_Paint_Mix_Act_Red_Tank_Temp" : Real = PLC Paramters_Paint_Mix.Act_Red_Tank_Temp, 1 s
   "Paramters_Paint_Mix_Act_Green_Tank_Temp" : Real = PLC Paramters_Paint_Mix.Act_Green_Tank_Temp, 1 s
   "Paramters_Paint_Mix_Act_Blue_Tank_Temp" : Real = PLC Paramters_Paint_Mix.Act_Blue_Tank_Temp, 1 s
   "Paramters_Paint_Mix_Act_Red_Tank_Press" : Real = PLC Paramters_Paint_Mix.Act_Red_Tank_Press, 1 s
   "Paramters_Paint_Mix_Act_Green_Tank_Press" : Real = PLC Paramters_Paint_Mix.Act_Green_Tank_Press, 1 s
   "Paramters_Paint_Mix_Act_Blue_Tank_Press" : Real = PLC Paramters_Paint_Mix.Act_Blue_Tank_Press, 1 s
   "PainMix_DB_Green_Tank_Level" : Int = PLC PainMix_DB.Green_Tank_Level, 1 s
   "PainMix_DB_Blue_Tank_Level" : Int = PLC PainMix_DB.Blue_Tank_Level, 1 s
   "PainMix_DB_Sol_1_Tank_Level" : Int = PLC PainMix_DB.Sol_1_Tank_Level, 1 s
   "PainMix_DB_Sol_2_Tank_Level" : Int = PLC PainMix_DB.Sol_2_Tank_Level, 1 s
   "Recipe_Pigment Concentration" : Real = PLC Recipe."Pigment Concentration", 1 s
   "Recipe_Resin Type and Ratio" : Real = PLC Recipe."Resin Type and Ratio", 1 s
   "Recipe_Solvent Composition" : Real = PLC Recipe."Solvent Composition", 1 s
   "Recipe_Additive Ratios" : Real = PLC Recipe."Additive Ratios", 1 s
   "Recipe_Drying Agent Ratio" : Real = PLC Recipe."Drying Agent Ratio", 1 s
   "Recipe_Viscosity Target" : Real = PLC Recipe."Viscosity Target", 1 s
   "Recipe_Gloss Level" : Real = PLC Recipe."Gloss Level", 1 s
   "Recipe_pH Control Range" : Real = PLC Recipe."pH Control Range", 1 s
   "Recipe_Mixing Time" : Real = PLC Recipe."Mixing Time", 1 s
   "Recipe_Curing Agent Proportion" : Real = PLC Recipe."Curing Agent Proportion", 1 s
   "Recipe_Recipe_Name" : String[254] = PLC Recipe.Recipe_Name, 1 s
   "PainMix_DB_MainTank_Mixer_Cont" : Bool = PLC PainMix_DB.MainTank_Mixer_Cont, 1 s
   "PainMix_DB_MainTank_Tank_Level" : Int = PLC PainMix_DB.MainTank_Tank_Level, 1 s
   "Paramters_Paint_Mix_Recipe_ID" : String[254] = PLC Paramters_Paint_Mix.Recipe_ID, 1 s
   "Paramters_Paint_Mix_Recipe_Name" : String[254] = PLC Paramters_Paint_Mix.Recipe_Name, 1 s
   "Paramters_Paint_Mix_Equip_ID" : String[254] = PLC Paramters_Paint_Mix.Equip_ID, 1 s
   "Paramters_Paint_Mix_Batch_ID" : String[254] = PLC Paramters_Paint_Mix.Batch_ID, 1 s
   "Paramters_Paint_Mix_Batch_Size" : String[254] = PLC Paramters_Paint_Mix.Batch_Size, 1 s
   "Paramters_Paint_Mix_Start_Time" : String[254] = PLC Paramters_Paint_Mix.Start_Time, 1 s
   "Paramters_Paint_Mix_Warning_1" : Bool = PLC Paramters_Paint_Mix.Warning_1, 1 s
   "Paramters_Paint_Mix_Warning_2" : Bool = PLC Paramters_Paint_Mix.Warning_2, 1 s
   "Paramters_Paint_Mix_Warning_3" : Bool = PLC Paramters_Paint_Mix.Warning_3, 1 s
   "Paramters_Paint_Mix_Alarm_1" : Bool = PLC Paramters_Paint_Mix.Alarm_1, 1 s
   "Paramters_Paint_Mix_Alarm_2" : Bool = PLC Paramters_Paint_Mix.Alarm_2, 1 s
   "Paramters_Paint_Mix_Common_A-W" : Bool = PLC Paramters_Paint_Mix.Common_A-W, 1 s
   "PainMix_DB_Alarm_ACK" : Bool = PLC PainMix_DB.Alarm_ACK, 1 s
   "Paramters_Paint_Mix_Language" : Bool = PLC Paramters_Paint_Mix.Language, 500 ms
   "Paramters_Paint_Mix_Button_Language" : Bool = PLC Paramters_Paint_Mix.Button_Language, 1 s
   "UserName_fromHMI" : WString[254] AT %DB1.DBD0
   "Paramters_Paint_Mix_MainOverview" : Bool = PLC Paramters_Paint_Mix.MainOverview, 1 s
   "Paramters_Paint_Mix_Parameters" : Bool = PLC Paramters_Paint_Mix.Parameters, 1 s
   "Paramters_Paint_Mix_RecipeM" : Bool = PLC Paramters_Paint_Mix.RecipeM, 1 s
   "Paramters_Paint_Mix_UserM" : Bool = PLC Paramters_Paint_Mix.UserM, 1 s
   "Paramters_Paint_Mix_AlarmSt" : Bool = PLC Paramters_Paint_Mix.AlarmSt, 1 s
   "Paramters_Paint_Mix_IOSt" : Bool = PLC Paramters_Paint_Mix.IOSt, 1 s

HMI tags "Paint_Mix"
   "MainT_Agitator" : Int = PLC PainMix_DB.Agitator_MainT, 500 ms

graphic list "Agitator": 0 'Graphic_92'; 1 'Graphic_91'; 2 'Graphic_93'

graphic list "Pump_Fan_Green": 0 'Graphic_67'; 1 'Graphic_68'; 2 'Graphic_69'; 3 'Graphic_70'

graphic list "Pump_Fan_Red": 0 'Graphic_80'; 1 'Graphic_81'; 2 'Graphic_82'; 3 'Graphic_83'

graphic list "Pump_Fan_Blue": 0 'Graphic_37'; 1 'Graphic_72'; 2 'Graphic_73'; 3 'Graphic_74'

recipe "Recipe_1": Recipe_element_1 <- "Recipe_Pigment Concentration", Recipe_element_2 <- "Recipe_Resin Type and Ratio", Recipe_element_3 <- "Recipe_Solvent Composition", Recipe_element_4 <- "Recipe_Additive Ratios", Recipe_element_5 <- "Recipe_Drying Agent Ratio", Recipe_element_6 <- "Recipe_Viscosity Target", Recipe_element_7 <- "Recipe_Gloss Level", Recipe_element_8 <- "Recipe_pH Control Range", Recipe_element_9 <- "Recipe_Mixing Time", Recipe_element_10 <- "Recipe_Curing Agent Proportion"

screen "MainOverview" 800x480, template "PaintMix"
   GraphicView "Graphic view_22" at 170,409 size 606x10; Picture "Graphic_48"
   GraphicView "Graphic view_33" at 755,401 size 18x18; Picture "Graphic_55"
   GraphicView "Graphic view_34" at 763,149 size 10x260; Picture "Graphic_54"
   GraphicView "Graphic view_35" at 755,142 size 18x18; Picture "Graphic_49"
   GraphicView "Graphic view_36" at 730,142 size 29x10; Picture "Graphic_48"
   GraphicView "Graphic view_29" at 714,142 size 18x18; Picture "Graphic_51"
   GraphicView "Graphic view_37" at 714,155 size 10x18; Picture "Graphic_54"
   GraphicView "Graphic view_23" at 187,233 size 18x18; Picture "Graphic_49"
   GraphicView "Graphic view_27" at 195,245 size 10x151; Picture "Graphic_54"
   GraphicView "Graphic view_24" at 195,386 size 18x18; Picture "Graphic_50"
   GraphicView "Graphic view_26" at 194,394 size 566x10; Picture "Graphic_48"
   GraphicView "Graphic view_32" at 741,386 size 18x18; Picture "Graphic_55"
   GraphicView "Graphic view_30" at 749,164 size 10x230; Picture "Graphic_54"
   GraphicView "Graphic view_31" at 741,155 size 18x18; Picture "Graphic_49"
   GraphicView "Graphic view_28" at 726,155 size 18x18; Picture "Graphic_51"
   GraphicView "Graphic view_47" at 355,235 size 10x73; Picture "Graphic_54"
   GraphicView "Graphic view_38" at 355,305 size 18x18; Picture "Graphic_50"
   GraphicView "Graphic view_44" at 365,313 size 126x10; Picture "Graphic_48"
   GraphicView "Graphic view_52" at 534,325 size 20x10; Picture "Graphic_48"
   GraphicView "Graphic view_51" at 551,317 size 18x18; Picture "Graphic_55"
   GraphicView "Graphic view_56" at 559,149 size 10x174; Picture "Graphic_54"
   GraphicView "Graphic view_61" at 559,142 size 18x18; Picture "Graphic_51"
   GraphicView "Graphic view_60" at 575,142 size 29x10; Picture "Graphic_48"
   GraphicView "Graphic view_62" at 600,142 size 18x18; Picture "Graphic_49"
   GraphicView "Graphic view_63" at 608,155 size 10x18; Picture "Graphic_54"
   GraphicView "Graphic view_48" at 457,234 size 10x36; Picture "Graphic_54"
   GraphicView "Graphic view_49" at 457,267 size 18x18; Picture "Graphic_50"
   GraphicView "Graphic view_50" at 473,275 size 14x10; Picture "Graphic_48"
   GraphicView "Graphic view_39" at 535,278 size 18x18; Picture "Graphic_55"
   GraphicView "Graphic view_55" at 543,131 size 10x155; Picture "Graphic_54"
   GraphicView "Graphic view_65" at 543,127 size 18x18; Picture "Graphic_51"
   GraphicView "Graphic view_64" at 558,127 size 61x10; Picture "Graphic_48"
   GraphicView "Graphic view_66" at 613,127 size 18x18; Picture "Graphic_49"
   GraphicView "Graphic view_67" at 621,139 size 10x35; Picture "Graphic_54"
   GraphicView "Graphic view_59" at 588,155 size 18x18; Picture "Graphic_49"
   GraphicView "Graphic view_58" at 573,155 size 18x18; Picture "Graphic_51"
   GraphicView "Graphic view_57" at 573,162 size 10x199; Picture "Graphic_54"
   GraphicView "Graphic view_54" at 565,354 size 18x18; Picture "Graphic_55"
   GraphicView "Graphic view_53" at 535,362 size 41x10; Picture "Graphic_48"
   GraphicView "Graphic view_41" at 292,352 size 202x10; Picture "Graphic_48"
   GraphicView "Graphic view_46" at 253,344 size 18x18; Picture "Graphic_50"
   GraphicView "Graphic view_40" at 253,235 size 10x115; Picture "Graphic_54"
   Rectangle "Rectangle_13" at 702,84 size 91x44
      Appearance <- "PainMix_DB_Control_Mode"
   GraphicView "Graphic view_43" at 122,409 size 34x10; Picture "Graphic_48"
   GraphicView "Graphic view_14" at 95,385 size 28x37; Picture "Graphic_46"
   GraphicView "Graphic view_17" at 95,209 size 28x37; Picture "Graphic_46"
   GraphicView "Graphic view_19" at 121,233 size 34x10; Picture "Graphic_48"
   TextField "Template_Text field_2" at 341,43 size 151x25; Text 'Hauptübersicht / Main Overview'
   GraphicView "Graphic view_2" at 586,166 size 158x222; Picture "Graphic_34"
   GraphicView "Graphic view_9" at 15,103 size 89x150; Picture "Graphic_22"
   GraphicView "Graphic view_10" at 206,80 size 103x141; Picture "Graphic_24"
   GraphicView "Graphic view_6" at 307,80 size 106x141; Picture "Graphic_24"
   GraphicView "Graphic view_12" at 411,80 size 103x141; Picture "Graphic_24"
   GraphicView "Graphic view_11" at 15,279 size 89x150; Picture "Graphic_22"
   GraphicView "Graphic view_13" at 351,206 size 44x34; Picture "Graphic_40"
   GraphicView "Graphic view_15" at 453,206 size 44x34; Picture "Graphic_40"
   GraphicView "Graphic view_16" at 249,206 size 44x34; Picture "Graphic_40"
   GraphicView "Graphic view_1" at 151,200 size 37x45; Picture "Graphic_39"
   Rectangle "Rectangle_2" at 102,387 size 14x13
      Appearance <- "PainMix_DB_Sol_2_Valve_Status"
   Bar "Bar_1" at 388,93 size 18x72; MinimumValue 0; MaximumValue 50
      ProcessValue <- "PainMix_DB_Green_Tank_Level"
   Bar "Bar_2" at 285,93 size 18x72; MinimumValue 0; MaximumValue 50
      ProcessValue <- "PainMix_DB_Red_Tank_Level"
   Bar "Bar_3" at 490,93 size 18x72; MinimumValue 0; MaximumValue 50
      ProcessValue <- "PainMix_DB_Blue_Tank_Level"
   Bar "Bar_4" at 45,130 size 28x94; MinimumValue 0; MaximumValue 50
      ProcessValue <- "PainMix_DB_Sol_1_Tank_Level"
   Bar "Bar_5" at 44,304 size 28x94; MinimumValue 0; MaximumValue 50
      ProcessValue <- "PainMix_DB_Sol_2_Tank_Level"
   GraphicView "Graphic view_7" at 268,314 size 33x54; Picture "Graphic_16"
   Bar "Bar_6" at 622,200 size 89x97; MinimumValue 0; MaximumValue 50
      ProcessValue <- "PainMix_DB_MainTank_Tank_Level"
   GraphicIOField "Graphic I/O field_1" at 649,196 size 37x105; PictureList "Agitator"
      ProcessValue <- "MainT_Agitator"
   GraphicView "Graphic view_45" at 485,272 size 51x37; Picture "Graphic_59"
   GraphicView "Graphic view_73" at 485,310 size 51x37; Picture "Graphic_59"
   GraphicView "Graphic view_42" at 485,348 size 51x37; Picture "Graphic_59"
   GraphicIOField "Graphic I/O field_2" at 499,278 size 27x27; PictureList "Pump_Fan_Blue"
      ProcessValue <- "PainMix_DB_Blue_P_Rotor"
   GraphicIOField "Graphic I/O field_3" at 499,316 size 27x27; PictureList "Pump_Fan_Green"
      ProcessValue <- "PainMix_DB_Green_P_Rotor"
   GraphicIOField "Graphic I/O field_4" at 499,354 size 27x27; PictureList "Pump_Fan_Red"
      ProcessValue <- "PainMix_DB_Red_P_Rotor"
   GraphicView "Graphic view_70" at 655,139 size 25x34; Picture "Graphic_95"
   Group "Group" at 170,142 size 606x277; Picture "Graphic_48"
   GraphicView "Graphic view_20" at 151,377 size 37x45; Picture "Graphic_39"
   Group "Group_1" at 187,155 size 573x249; Picture "Graphic_49"
   IOField "Template_I/O field_1" at 218,109 size 58x17; FormatPattern 99.9; Unit  °C
      ProcessValue <- "Paramters_Paint_Mix_Act_Red_Tank_Temp"
   TextField "Template_Text field_1" at 206,94 size 82x15; Text 'Temperatur / Temperature'
   IOField "Template_I/O field_2" at 218,142 size 58x17; FormatPattern 99.9; Unit  bar
      ProcessValue <- "Paramters_Paint_Mix_Act_Red_Tank_Press"
   TextField "Template_Text field_3" at 218,128 size 58x15; Text 'Druck / Pressure'
   GraphicView "Graphic view_71" at 194,249 size 13x30; Picture "Graphic_99"
      Visibility <- "PainMix_DB_Sol_1_Pipe1"
   GraphicView "Graphic view_79" at 122,232 size 31x13; Picture "Graphic_104"
      Visibility <- "PainMix_DB_Sol_1_Pipe1"
   GraphicView "Graphic view_80" at 210,393 size 30x13; Picture "Graphic_104"
      Visibility <- "PainMix_DB_Sol_1_Pipe1"
   GraphicView "Graphic view_81" at 194,276 size 13x30; Picture "Graphic_99"
      Visibility <- "PainMix_DB_Sol_1_Pipe1"
   GraphicView "Graphic view_82" at 194,303 size 13x30; Picture "Graphic_99"
      Visibility <- "PainMix_DB_Sol_1_Pipe1"
   GraphicView "Graphic view_83" at 194,330 size 13x30; Picture "Graphic_99"
      Visibility <- "PainMix_DB_Sol_1_Pipe1"
   GraphicView "Graphic view_84" at 194,357 size 13x33; Picture "Graphic_99"
      Visibility <- "PainMix_DB_Sol_1_Pipe1"
   GraphicView "Graphic view_78" at 238,393 size 30x13; Picture "Graphic_104"
      Visibility <- "PainMix_DB_Sol_1_Pipe1"
   GraphicView "Graphic view_85" at 266,393 size 30x13; Picture "Graphic_104"
      Visibility <- "PainMix_DB_Sol_1_Pipe1"
   GraphicView "Graphic view_86" at 294,393 size 30x13; Picture "Graphic_104"
      Visibility <- "PainMix_DB_Sol_1_Pipe1"
   GraphicView "Graphic view_87" at 322,393 size 30x13; Picture "Graphic_104"
      Visibility <- "PainMix_DB_Sol_1_Pipe1"
   GraphicView "Graphic view_88" at 350,393 size 30x13; Picture "Graphic_104"
      Visibility <- "PainMix_DB_Sol_1_Pipe1"
   GraphicView "Graphic view_89" at 378,393 size 30x13; Picture "Graphic_104"
      Visibility <- "PainMix_DB_Sol_1_Pipe1"
   GraphicView "Graphic view_90" at 406,393 size 30x13; Picture "Graphic_104"
      Visibility <- "PainMix_DB_Sol_1_Pipe1"
   GraphicView "Graphic view_91" at 434,393 size 30x13; Picture "Graphic_104"
      Visibility <- "PainMix_DB_Sol_1_Pipe1"
   GraphicView "Graphic view_92" at 462,393 size 30x13; Picture "Graphic_104"
      Visibility <- "PainMix_DB_Sol_1_Pipe1"
   GraphicView "Graphic view_93" at 490,393 size 30x13; Picture "Graphic_104"
      Visibility <- "PainMix_DB_Sol_1_Pipe1"
   GraphicView "Graphic view_94" at 518,393 size 30x13; Picture "Graphic_104"
      Visibility <- "PainMix_DB_Sol_1_Pipe1"
   GraphicView "Graphic view_95" at 546,393 size 30x13; Picture "Graphic_104"
      Visibility <- "PainMix_DB_Sol_1_Pipe1"
   GraphicView "Graphic view_96" at 574,393 size 30x13; Picture "Graphic_104"
      Visibility <- "PainMix_DB_Sol_1_Pipe1"
   GraphicView "Graphic view_97" at 602,393 size 30x13; Picture "Graphic_104"
      Visibility <- "PainMix_DB_Sol_1_Pipe1"
   GraphicView "Graphic view_98" at 630,393 size 30x13; Picture "Graphic_104"
      Visibility <- "PainMix_DB_Sol_1_Pipe1"
   GraphicView "Graphic view_99" at 658,393 size 30x13; Picture "Graphic_104"
      Visibility <- "PainMix_DB_Sol_1_Pipe1"
   GraphicView "Graphic view_100" at 686,393 size 30x13; Picture "Graphic_104"
      Visibility <- "PainMix_DB_Sol_1_Pipe1"
   GraphicView "Graphic view_101" at 714,393 size 30x13; Picture "Graphic_104"
      Visibility <- "PainMix_DB_Sol_1_Pipe1"
   GraphicView "Graphic view_102" at 748,248 size 13x30; Picture "Graphic_99"
      Visibility <- "PainMix_DB_Sol_1_Pipe1"
   GraphicView "Graphic view_103" at 748,275 size 13x30; Picture "Graphic_99"
      Visibility <- "PainMix_DB_Sol_1_Pipe1"
   GraphicView "Graphic view_104" at 748,302 size 13x30; Picture "Graphic_99"
      Visibility <- "PainMix_DB_Sol_1_Pipe1"
   GraphicView "Graphic view_105" at 748,329 size 13x30; Picture "Graphic_99"
      Visibility <- "PainMix_DB_Sol_1_Pipe1"
   GraphicView "Graphic view_106" at 748,356 size 13x33; Picture "Graphic_99"
      Visibility <- "PainMix_DB_Sol_1_Pipe1"
   GraphicView "Graphic view_107" at 748,166 size 13x31; Picture "Graphic_99"
      Visibility <- "PainMix_DB_Sol_1_Pipe1"
   GraphicView "Graphic view_108" at 748,194 size 13x30; Picture "Graphic_99"
      Visibility <- "PainMix_DB_Sol_1_Pipe1"
   GraphicView "Graphic view_109" at 748,221 size 13x30; Picture "Graphic_99"
      Visibility <- "PainMix_DB_Sol_1_Pipe1"
   GraphicView "Graphic view_110" at 725,166 size 13x8; Picture "Graphic_99"
      Visibility <- "PainMix_DB_Sol_1_Pipe1"
   GraphicView "Graphic view_111" at 187,408 size 30x13; Picture "Graphic_105"
      Visibility <- "PainMix_DB_Sol_1_Pipe2"
   GraphicView "Graphic view_112" at 215,408 size 30x13; Picture "Graphic_105"
      Visibility <- "PainMix_DB_Sol_1_Pipe2"
   GraphicView "Graphic view_113" at 243,408 size 30x13; Picture "Graphic_105"
      Visibility <- "PainMix_DB_Sol_1_Pipe2"
   GraphicView "Graphic view_114" at 271,408 size 30x13; Picture "Graphic_105"
      Visibility <- "PainMix_DB_Sol_1_Pipe2"
   GraphicView "Graphic view_115" at 299,408 size 30x13; Picture "Graphic_105"
      Visibility <- "PainMix_DB_Sol_1_Pipe2"
   GraphicView "Graphic view_116" at 327,408 size 30x13; Picture "Graphic_105"
      Visibility <- "PainMix_DB_Sol_1_Pipe2"
   GraphicView "Graphic view_117" at 355,408 size 30x13; Picture "Graphic_105"
      Visibility <- "PainMix_DB_Sol_1_Pipe2"
   GraphicView "Graphic view_118" at 383,408 size 30x13; Picture "Graphic_105"
      Visibility <- "PainMix_DB_Sol_1_Pipe2"
   GraphicView "Graphic view_119" at 411,408 size 30x13; Picture "Graphic_105"
      Visibility <- "PainMix_DB_Sol_1_Pipe2"
   GraphicView "Graphic view_120" at 439,408 size 30x13; Picture "Graphic_105"
      Visibility <- "PainMix_DB_Sol_1_Pipe2"
   GraphicView "Graphic view_121" at 467,408 size 30x13; Picture "Graphic_105"
      Visibility <- "PainMix_DB_Sol_1_Pipe2"
   GraphicView "Graphic view_122" at 495,408 size 30x13; Picture "Graphic_105"
      Visibility <- "PainMix_DB_Sol_1_Pipe2"
   GraphicView "Graphic view_123" at 523,408 size 30x13; Picture "Graphic_105"
      Visibility <- "PainMix_DB_Sol_1_Pipe2"
   GraphicView "Graphic view_124" at 551,408 size 30x13; Picture "Graphic_105"
      Visibility <- "PainMix_DB_Sol_1_Pipe2"
   GraphicView "Graphic view_125" at 579,408 size 30x13; Picture "Graphic_105"
      Visibility <- "PainMix_DB_Sol_1_Pipe2"
   GraphicView "Graphic view_126" at 607,408 size 30x13; Picture "Graphic_105"
      Visibility <- "PainMix_DB_Sol_1_Pipe2"
   GraphicView "Graphic view_127" at 635,408 size 30x13; Picture "Graphic_105"
      Visibility <- "PainMix_DB_Sol_1_Pipe2"
   GraphicView "Graphic view_128" at 663,408 size 30x13; Picture "Graphic_105"
      Visibility <- "PainMix_DB_Sol_1_Pipe2"
   GraphicView "Graphic view_129" at 691,408 size 30x13; Picture "Graphic_105"
      Visibility <- "PainMix_DB_Sol_1_Pipe2"
   GraphicView "Graphic view_130" at 123,408 size 30x13; Picture "Graphic_105"
      Visibility <- "PainMix_DB_Sol_1_Pipe2"
   GraphicView "Graphic view_132" at 762,239 size 13x30; Picture "Graphic_106"
      Visibility <- "PainMix_DB_Sol_1_Pipe2"
   GraphicView "Graphic view_133" at 762,266 size 13x30; Picture "Graphic_106"
      Visibility <- "PainMix_DB_Sol_1_Pipe2"
   GraphicView "Graphic view_134" at 762,293 size 13x30; Picture "Graphic_106"
      Visibility <- "PainMix_DB_Sol_1_Pipe2"
   GraphicView "Graphic view_135" at 762,320 size 13x30; Picture "Graphic_106"
      Visibility <- "PainMix_DB_Sol_1_Pipe2"
   GraphicView "Graphic view_136" at 762,347 size 13x33; Picture "Graphic_106"
      Visibility <- "PainMix_DB_Sol_1_Pipe2"
   GraphicView "Graphic view_137" at 762,157 size 13x31; Picture "Graphic_106"
      Visibility <- "PainMix_DB_Sol_1_Pipe2"
   GraphicView "Graphic view_138" at 762,185 size 13x30; Picture "Graphic_106"
      Visibility <- "PainMix_DB_Sol_1_Pipe2"
   GraphicView "Graphic view_139" at 762,212 size 13x30; Picture "Graphic_106"
      Visibility <- "PainMix_DB_Sol_1_Pipe2"
   GraphicView "Graphic view_140" at 762,378 size 13x26; Picture "Graphic_106"
      Visibility <- "PainMix_DB_Sol_1_Pipe2"
   GraphicView "Graphic view_141" at 720,408 size 38x13; Picture "Graphic_105"
      Visibility <- "PainMix_DB_Sol_1_Pipe2"
   GraphicView "Graphic view_144" at 729,141 size 33x13; Picture "Graphic_105"
      Visibility <- "PainMix_DB_Sol_1_Pipe2"
   GraphicView "Graphic view_145" at 713,156 size 13x18; Picture "Graphic_106"
      Visibility <- "PainMix_DB_Sol_1_Pipe2"
   Group "Group_2" at 253,155 size 353x217; Picture "Graphic_49"
   GraphicView "Graphic view_152" at 572,243 size 13x30; Picture "Graphic_108"
      Visibility <- "PainMix_DB_RED_Pipe"
   GraphicView "Graphic view_160" at 572,270 size 13x30; Picture "Graphic_108"
      Visibility <- "PainMix_DB_RED_Pipe"
   GraphicView "Graphic view_161" at 572,297 size 13x30; Picture "Graphic_108"
      Visibility <- "PainMix_DB_RED_Pipe"
   GraphicView "Graphic view_162" at 572,324 size 13x33; Picture "Graphic_108"
      Visibility <- "PainMix_DB_RED_Pipe"
   GraphicView "Graphic view_164" at 572,167 size 13x21; Picture "Graphic_108"
      Visibility <- "PainMix_DB_RED_Pipe"
   GraphicView "Graphic view_165" at 572,185 size 13x30; Picture "Graphic_108"
      Visibility <- "PainMix_DB_RED_Pipe"
   GraphicView "Graphic view_166" at 572,212 size 13x33; Picture "Graphic_108"
      Visibility <- "PainMix_DB_RED_Pipe"
   GraphicView "Graphic view_163" at 595,165 size 13x9; Picture "Graphic_108"
      Visibility <- "PainMix_DB_RED_Pipe"
   GraphicView "Graphic view_153" at 300,351 size 19x13; Picture "Graphic_107"
      Visibility <- "PainMix_DB_RED_Pipe"
   GraphicView "Graphic view_154" at 317,351 size 30x13; Picture "Graphic_107"
      Visibility <- "PainMix_DB_RED_Pipe"
   GraphicView "Graphic view_155" at 345,351 size 30x13; Picture "Graphic_107"
      Visibility <- "PainMix_DB_RED_Pipe"
   GraphicView "Graphic view_156" at 373,351 size 30x13; Picture "Graphic_107"
      Visibility <- "PainMix_DB_RED_Pipe"
   GraphicView "Graphic view_157" at 401,351 size 30x13; Picture "Graphic_107"
      Visibility <- "PainMix_DB_RED_Pipe"
   GraphicView "Graphic view_158" at 429,351 size 30x13; Picture "Graphic_107"
      Visibility <- "PainMix_DB_RED_Pipe"
   GraphicView "Graphic view_159" at 457,351 size 32x13; Picture "Graphic_107"
      Visibility <- "PainMix_DB_RED_Pipe"
   GraphicView "Graphic view_147" at 252,314 size 13x34; Picture "Graphic_108"
      Visibility <- "PainMix_DB_RED_Pipe"
   GraphicView "Graphic view_167" at 252,237 size 13x22; Picture "Graphic_108"
      Visibility <- "PainMix_DB_RED_Pipe"
   GraphicView "Graphic view_168" at 252,256 size 13x30; Picture "Graphic_108"
      Visibility <- "PainMix_DB_RED_Pipe"
   GraphicView "Graphic view_169" at 252,283 size 13x33; Picture "Graphic_108"
      Visibility <- "PainMix_DB_RED_Pipe"
   GraphicView "Graphic view_148" at 536,361 size 35x13; Picture "Graphic_107"
      Visibility <- "PainMix_DB_RED_Pipe"
   Group "Group_3" at 355,142 size 263x193; Picture "Graphic_54"
   GraphicView "Graphic view_68" at 373,275 size 33x54; Picture "Graphic_16"
   Group "Group_4" at 457,127 size 174x169; Picture "Graphic_54"
   GraphicView "Graphic view_69" at 573,93 size 30x49; Picture "Graphic_16"
   GraphicView "Graphic view_150" at 354,237 size 13x22; Picture "Graphic_99"
      Visibility <- "PainMix_DB_GREEN_Pipe"
   GraphicView "Graphic view_151" at 354,256 size 13x30; Picture "Graphic_99"
      Visibility <- "PainMix_DB_GREEN_Pipe"
   GraphicView "Graphic view_170" at 354,283 size 13x24; Picture "Graphic_99"
      Visibility <- "PainMix_DB_GREEN_Pipe"
   GraphicView "Graphic view_149" at 558,249 size 13x22; Picture "Graphic_99"
      Visibility <- "PainMix_DB_GREEN_Pipe"
   GraphicView "Graphic view_171" at 558,268 size 13x30; Picture "Graphic_99"
      Visibility <- "PainMix_DB_GREEN_Pipe"
   GraphicView "Graphic view_172" at 558,295 size 13x24; Picture "Graphic_99"
      Visibility <- "PainMix_DB_GREEN_Pipe"
   GraphicView "Graphic view_173" at 558,182 size 13x22; Picture "Graphic_99"
      Visibility <- "PainMix_DB_GREEN_Pipe"
   GraphicView "Graphic view_174" at 558,201 size 13x30; Picture "Graphic_99"
      Visibility <- "PainMix_DB_GREEN_Pipe"
   GraphicView "Graphic view_175" at 558,228 size 13x24; Picture "Graphic_99"
      Visibility <- "PainMix_DB_GREEN_Pipe"
   GraphicView "Graphic view_177" at 558,156 size 13x16; Picture "Graphic_99"
      Visibility <- "PainMix_DB_GREEN_Pipe"
   GraphicView "Graphic view_178" at 558,169 size 13x16; Picture "Graphic_99"
      Visibility <- "PainMix_DB_GREEN_Pipe"
   GraphicView "Graphic view_176" at 606,155 size 15x19; Picture "Graphic_99"
      Visibility <- "PainMix_DB_GREEN_Pipe"
   GraphicView "Graphic view_179" at 404,312 size 26x13; Picture "Graphic_104"
      Visibility <- "PainMix_DB_GREEN_Pipe"
   GraphicView "Graphic view_180" at 428,312 size 30x13; Picture "Graphic_104"
      Visibility <- "PainMix_DB_GREEN_Pipe"
   GraphicView "Graphic view_181" at 456,312 size 32x13; Picture "Graphic_104"
      Visibility <- "PainMix_DB_GREEN_Pipe"
   GraphicView "Graphic view_182" at 575,141 size 29x13; Picture "Graphic_104"
      Visibility <- "PainMix_DB_GREEN_Pipe"
   GraphicView "Graphic view_185" at 542,210 size 13x22; Picture "Graphic_109"
      Visibility <- "PainMix_DB_BLUE_Pipe"
   GraphicView "Graphic view_186" at 542,229 size 13x30; Picture "Graphic_109"
      Visibility <- "PainMix_DB_BLUE_Pipe"
   GraphicView "Graphic view_187" at 542,256 size 13x24; Picture "Graphic_109"
      Visibility <- "PainMix_DB_BLUE_Pipe"
   GraphicView "Graphic view_188" at 542,143 size 13x22; Picture "Graphic_109"
      Visibility <- "PainMix_DB_BLUE_Pipe"
   GraphicView "Graphic view_189" at 542,162 size 13x30; Picture "Graphic_109"
      Visibility <- "PainMix_DB_BLUE_Pipe"
   GraphicView "Graphic view_190" at 542,189 size 13x24; Picture "Graphic_109"
      Visibility <- "PainMix_DB_BLUE_Pipe"
   GraphicView "Graphic view_191" at 558,126 size 17x13; Picture "Graphic_110"
      Visibility <- "PainMix_DB_BLUE_Pipe"
   GraphicView "Graphic view_192" at 602,126 size 16x13; Picture "Graphic_110"
      Visibility <- "PainMix_DB_BLUE_Pipe"
   GraphicView "Graphic view_74" at 456,236 size 13x21; Picture "Graphic_109"
      Visibility <- "PainMix_DB_BLUE_Pipe"
   GraphicView "Graphic view_75" at 456,254 size 13x20; Picture "Graphic_109"
      Visibility <- "PainMix_DB_BLUE_Pipe"
   GraphicView "Graphic view_76" at 620,140 size 13x22; Picture "Graphic_109"
      Visibility <- "PainMix_DB_BLUE_Pipe"
   GraphicView "Graphic view_77" at 620,159 size 13x15; Picture "Graphic_109"
      Visibility <- "PainMix_DB_BLUE_Pipe"
   GraphicView "Graphic view_131" at 535,324 size 22x13; Picture "Graphic_104"
      Visibility <- "PainMix_DB_GREEN_Pipe"
   GraphicView "Graphic view_142" at 471,274 size 17x13; Picture "Graphic_110"
      Visibility <- "PainMix_DB_BLUE_Pipe"
   TextField "Template_Text field_9" at 4,79 size 110x30; Text 'Harzverst. Tank Resin Enhancer Tank'
   TextField "Template_Text field_10" at 210,169 size 95x26; Text 'Rot Pigm. Tank RED Pigment Tank'
   TextField "Template_Text field_11" at 308,169 size 103x26; Text 'Grün Pigm. Tank GREEN Pigment Tank'
   TextField "Template_Text field_12" at 412,169 size 101x26; Text 'Blau Pigm. Tank BLUE Pigment Tank'
   Rectangle "Rectangle_6" at 162,374 size 15x10
      Appearance <- "PainMix_DB_Sol_2_Valve_Status"
   Rectangle "Rectangle_7" at 102,211 size 14x13
      Appearance <- "PainMix_DB_Sol_1_Valve_Status"
   Rectangle "Rectangle_8" at 162,197 size 15x10
      Appearance <- "PainMix_DB_Sol_1_Valve_Status"
   TextField "Template_Text field_13" at 615,176 size 103x18; Text 'Mischbehälter / Mixing Tank'
   Rectangle "Rectangle_1" at 657,143 size 22x13
      Appearance <- "PainMix_DB_MainTank_Mixer_Status"
   Rectangle "Rectangle_9" at 282,217 size 10x19
      Appearance <- "PainMix_DB_Red_Valve_Status"
   Rectangle "Rectangle_10" at 384,217 size 10x19
      Appearance <- "PainMix_DB_Green_Valve_Status"
   Rectangle "Rectangle_11" at 486,217 size 10x19
      Appearance <- "PainMix_DB_Blue_Valve_Status"
   GraphicView "Graphic view_3" at 123,208 size 23x23; Picture "tap_1196455"
      Visibility <- "PainMix_DB_Control_Mode"
   GraphicView "Graphic view_4" at 123,383 size 23x23; Picture "tap_1196455"
      Visibility <- "PainMix_DB_Control_Mode"
   GraphicView "Graphic view_5" at 296,225 size 23x23; Picture "tap_1196455"
      Visibility <- "PainMix_DB_Control_Mode"
   GraphicView "Graphic view_8" at 398,225 size 23x23; Picture "tap_1196455"
      Visibility <- "PainMix_DB_Control_Mode"
   GraphicView "Graphic view_18" at 500,225 size 23x23; Picture "tap_1196455"
      Visibility <- "PainMix_DB_Control_Mode"
   GraphicView "Graphic view_21" at 681,143 size 23x23; Picture "tap_1196455"
      Visibility <- "PainMix_DB_Control_Mode"
   Button "Button_1" at 102,209 size 45x20; TextOff 'Text'; Authorization "Operate"
      on Click: function_efd93a16("Resin_Valve_popup", 312, 166, -1, -1, 1)
      Visibility <- "PainMix_DB_Control_Mode"
   Button "Button_2" at 102,385 size 45x20; TextOff 'Text'; Authorization "Operate"
      Visibility <- "PainMix_DB_Control_Mode"
      on Click: function_efd93a16("Binder_Valve_popup", 312, 166, -1, -1, 1)
   Button "Button_3" at 270,217 size 51x29; TextOff 'Text'; Authorization "Operate"
      Visibility <- "PainMix_DB_Control_Mode"
      on Click: function_efd93a16("Red_Valve_popup", 312, 166, -1, -1, 1)
   Button "Button_4" at 371,217 size 51x29; TextOff 'Text'; Authorization "Operate"
      Visibility <- "PainMix_DB_Control_Mode"
      on Click: function_efd93a16("Green_Valve_popup", 312, 166, -1, -1, 1)
   Button "Button_5" at 472,217 size 51x29; TextOff 'Text'; Authorization "Operate"
      Visibility <- "PainMix_DB_Control_Mode"
      on Click: function_efd93a16("Blue_Valve_popup", 312, 166, -1, -1, 1)
   Button "Button_6" at 653,137 size 51x29; TextOff 'Text'; Authorization "Operate"
      Visibility <- "PainMix_DB_Control_Mode"
      on Click: function_efd93a16("MainTank_Valve_popup", 312, 166, -1, -1, 1)
   IOField "Template_I/O field_3" at 319,109 size 58x17; FormatPattern 99.9; Unit  °C
      ProcessValue <- "Paramters_Paint_Mix_Act_Green_Tank_Temp"
   TextField "Template_Text field_4" at 307,94 size 82x15; Text 'Temperatur / Temperature'
   IOField "Template_I/O field_4" at 319,142 size 58x17; FormatPattern 99.9; Unit  bar
      ProcessValue <- "Paramters_Paint_Mix_Act_Green_Tank_Press"
   TextField "Template_Text field_5" at 319,128 size 58x15; Text 'Druck / Pressure'
   IOField "Template_I/O field_5" at 423,109 size 58x17; FormatPattern 99.9; Unit  °C
      ProcessValue <- "Paramters_Paint_Mix_Act_Blue_Tank_Temp"
   TextField "Template_Text field_6" at 411,94 size 82x15; Text 'Temperatur / Temperature'
   IOField "Template_I/O field_6" at 423,142 size 58x17; FormatPattern 99.9; Unit  bar
      ProcessValue <- "Paramters_Paint_Mix_Act_Blue_Tank_Press"
   TextField "Template_Text field_7" at 423,128 size 58x15; Text 'Druck / Pressure'
   TextField "Template_Text field_17" at 4,253 size 110x30; Text 'Harzverst. Tank Solvent Binder Tank'
   Button "Button_7" at 696,84 size 103x46; TextOff 'Text'; Authorization "Operate"
      on Click: function_efd93a16("BatchDetails", 186, 74, -1, -1, 1)
   Button "Button_8" at 702,84 size 91x23; TextOff 'Control Panel / AN'; Authorization "Operate"
      on Click: function_efd93a16("BatchDetails", 186, 74, -1, -1, 1)
   TextField "Template_Text field_8" at 716,100 size 64x34; Text 'Lösungsmittelbinder / MANUAL'
      Visibility <- "PainMix_DB_Control_Mode"
   TextField "Template_Text field_14" at 716,100 size 64x34; Text 'Lösungsmittelbinder / AUTO'
      Visibility <- "PainMix_DB_Control_Mode"

Template "PaintMix" 800x480
   Button "Template_Button_7" at 0,1 size 799x80; TextOff 'Text'
   Button "Template_Button_1" at 0,434 size 111x44; TextOff 'Hauptübersicht Main Overview'; TextOn 'Main Overview Hauptübersicht'; Authorization "Monitor"
      on Click: ActivateScreen("MainOverview", 0); SetBit("Paramters_Paint_Mix_MainOverview"); ResetBit("Paramters_Paint_Mix_Parameters"); ResetBit("Paramters_Paint_Mix_RecipeM"); ResetBit("Paramters_Paint_Mix_UserM"); ResetBit("Paramters_Paint_Mix_AlarmSt"); ResetBit("Paramters_Paint_Mix_IOSt")
      Appearance <- "Paramters_Paint_Mix_MainOverview"
   Button "Template_Button_2" at 112,434 size 111x44; TextOn 'Parameter'; TextOff 'Parameter'; Authorization "Operate"
      on Click: ActivateScreen("Parameter", 0); SetBit("Paramters_Paint_Mix_Parameters"); ResetBit("Paramters_Paint_Mix_MainOverview"); ResetBit("Paramters_Paint_Mix_RecipeM"); ResetBit("Paramters_Paint_Mix_UserM"); ResetBit("Paramters_Paint_Mix_AlarmSt"); ResetBit("Paramters_Paint_Mix_IOSt")
      Appearance <- "Paramters_Paint_Mix_Parameters"
   Button "Template_Button_3" at 224,434 size 111x44; TextOn 'Recipe Management Rezept Verw.'; TextOff 'Rezept Verw. Recipe Management'; Authorization "User administration"
      on Click: ActivateScreen("Recipe", 0); SetBit("Paramters_Paint_Mix_RecipeM"); ResetBit("Paramters_Paint_Mix_Parameters"); ResetBit("Paramters_Paint_Mix_MainOverview"); ResetBit("Paramters_Paint_Mix_UserM"); ResetBit("Paramters_Paint_Mix_AlarmSt"); ResetBit("Paramters_Paint_Mix_IOSt")
      Appearance <- "Paramters_Paint_Mix_RecipeM"
   Button "Template_Button_4" at 336,434 size 111x44; TextOn 'User Management Ben. Verw.'; TextOff 'Ben. Verw. User Management'; Authorization "Monitor"
      on Click: ActivateScreen("User_Admin", 0); SetBit("Paramters_Paint_Mix_UserM"); ResetBit("Paramters_Paint_Mix_Parameters"); ResetBit("Paramters_Paint_Mix_RecipeM"); ResetBit("Paramters_Paint_Mix_MainOverview"); ResetBit("Paramters_Paint_Mix_AlarmSt"); ResetBit("Paramters_Paint_Mix_IOSt")
      Appearance <- "Paramters_Paint_Mix_UserM"
   Button "Template_Button_5" at 448,434 size 111x44; TextOn 'Alarm Status Alarm Status'; TextOff 'Alarm Status Alarm Status'; Authorization "Monitor"
      on Click: ActivateScreen("Alarm", 0); SetBit("Paramters_Paint_Mix_AlarmSt"); ResetBit("Paramters_Paint_Mix_Parameters"); ResetBit("Paramters_Paint_Mix_RecipeM"); ResetBit("Paramters_Paint_Mix_UserM"); ResetBit("Paramters_Paint_Mix_MainOverview"); ResetBit("Paramters_Paint_Mix_IOSt")
      Appearance <- "Paramters_Paint_Mix_AlarmSt"
   Button "Template_Button_6" at 560,434 size 111x44; TextOn 'I/O Status E/A-Status'; TextOff 'E/A-Status I/O Status'; Authorization "Monitor"
      on Click: ActivateScreen("Input_Status", 0); SetBit("Paramters_Paint_Mix_IOSt"); ResetBit("Paramters_Paint_Mix_Parameters"); ResetBit("Paramters_Paint_Mix_RecipeM"); ResetBit("Paramters_Paint_Mix_UserM"); ResetBit("Paramters_Paint_Mix_AlarmSt"); ResetBit("Paramters_Paint_Mix_MainOverview")
   GraphicView "Template_Graphic view_2" at 743,427 size 56x52; Picture "screenshot"
   Button "Template_Button_10" at 714,1 size 82x80; TextOff 'Text'
   Button "Template_Button_11" at 3,1 size 82x80; TextOff 'Text'
   GraphicView "Template_Graphic view_1" at 9,5 size 71x72; Picture "Dalle_1"
   Button "Template_Button_12" at 88,5 size 625x31; TextOff 'Text'
   DateTimeField "Template_Date/time field_1" at 87,37 size 107x38
   DateTimeField "Template_Date/time field_2" at 623,38 size 89x38
   Button "Template_Button_13" at 196,41 size 425x31; TextOff 'Text'
   TextField "Template_Text field_2" at 264,6 size 273x25; Text 'Farbherstellungsstation / Paint Manufacturing Station'
   TextField "Template_Text field_1" at 716,56 size 79x21; Text 'Nutzer / Username'
   IOField "Template_I/O field_1" at 717,33 size 78x24; FormatPattern ???????????????????????????????????????????????????????????????????
      ProcessValue <- "UserName_fromHMI"
   GraphicView "Template_Graphic view_3" at 734,0 size 40x33; Picture "Graphic_4"
   Button "Button_3" at 745,424 size 53x55; TextOff 'Text'
      on Click: function_f98d16b7()
   GraphicView "Graphic view_1" at 659,5 size 53x30; Picture "Graphic_114"
      Visibility <- "Paramters_Paint_Mix_Language"
   GraphicView "Graphic view_2" at 659,5 size 53x30; Picture "Graphic_116"
      Visibility <- "Paramters_Paint_Mix_Language"
   Button "Button_7" at 650,3 size 65x37; TextOff 'Text'
      on Click: function_fb9197e8(-1)
      on Release: ResetBit("Paramters_Paint_Mix_Button_Language")
      on Press: SetBit("Paramters_Paint_Mix_Button_Language")
   GraphicView "Template_Graphic view_4" at 522,411 size 43x43; Picture "Graphic_125"
      Visibility <- "Paramters_Paint_Mix_Common_A-W"

screen "Parameter" 800x480, template "PaintMix"
   TextField "Template_Text field_2" at 353,41 size 112x25; Text 'Parameter / Parameters'
   TextField "Template_Text field_9" at 6,85 size 144x23; Text 'Harzverstärker / Resin Enhancer'
   TextField "Template_Text field_1" at 13,111 size 133x20; Text 'Ausgangsfluss / Output Flow Rate'
   IOField "Template_I/O field_1" at 39,152 size 80x23; FormatPattern 99.9; Unit  m³/h
      ProcessValue <- "Paramters_Paint_Mix_ResinE_Flow_Act"
   TextField "Template_Text field_3" at 54,134 size 55x18; Text 'Aktuell / Actual'
   TextField "Template_Text field_4" at 46,178 size 67x18; Text 'Sollwert / Setpoint'
   IOField "Template_I/O field_2" at 44,196 size 80x23; FormatPattern 99.9; Unit  m³/h
      ProcessValue <- "Paramters_Paint_Mix_ResinE_Flow_Set"
   TextField "Template_Text field_5" at 4,228 size 147x18; Text 'Entsch. Sollw. / Defoaming Setpoint'
   IOField "Template_I/O field_3" at 43,248 size 71x23; FormatPattern 99.9; Unit  %
      ProcessValue <- "Paramters_Paint_Mix_Defoaming_Set"
   TextField "Template_Text field_6" at 164,112 size 133x20; Text 'Ausgangsfluss / Output Flow Rate'
   IOField "Template_I/O field_4" at 190,153 size 80x23; FormatPattern 99.9; Unit  m³/h
      ProcessValue <- "Paramters_Paint_Mix_Binder_Flow_Act"
   TextField "Template_Text field_7" at 205,135 size 55x18; Text 'Aktuell / Actual'
   TextField "Template_Text field_8" at 197,179 size 67x18; Text 'Sollwert / Setpoint'
   IOField "Template_I/O field_5" at 190,197 size 80x23; FormatPattern 99.9; Unit  m³/h
      ProcessValue <- "Paramters_Paint_Mix_Binder_Flow_Set"
   TextField "Template_Text field_10" at 156,229 size 151x18; Text 'Glanzverh.-Sollw. / Gloss Ratio Setpoint'
   IOField "Template_I/O field_6" at 194,249 size 71x23; FormatPattern 99.9; Unit  %
      ProcessValue <- "Paramters_Paint_Mix_Gloss Ratio_Set"
   TextField "Template_Text field_11" at 134,85 size 190x23; Text 'Lösungsmittelbinder / Solvent Binder'
   TextField "Template_Text field_15" at 318,85 size 138x23; Text 'Rotes Pigment / RED Pigment'
   TextField "Template_Text field_12" at 331,115 size 108x18; Text 'Füllst.-Sollw. / Level Setpoint'
   IOField "Template_I/O field_7" at 350,135 size 71x23; FormatPattern 99.9; Unit  ltr
      ProcessValue <- "Paramters_Paint_Mix_Level_Set_R"
   TextField "Template_Text field_13" at 319,166 size 133x18; Text 'Durchfluss-Sollw. / Flowrate Setpoint'
   IOField "Template_I/O field_8" at 345,186 size 80x23; FormatPattern 99.9; Unit  m³/h
      ProcessValue <- "Paramters_Paint_Mix_Flowrate_Set_R"
   TextField "Template_Text field_14" at 318,218 size 147x18; Text 'Viskositäts-Sollwert / Viscosity Setpoint'
   IOField "Template_I/O field_9" at 350,238 size 71x23; FormatPattern 99.9; Unit  cP
      ProcessValue <- "Paramters_Paint_Mix_Viscosity_Set_R"
   TextField "Template_Text field_16" at 305,320 size 161x18; Text 'Temp.-Sollwert / Temperature Setpoint'
   IOField "Template_I/O field_10" at 350,339 size 71x23; FormatPattern 99.9; Unit  °C
      ProcessValue <- "Paramters_Paint_Mix_Temperature_Set_R"
   TextField "Template_Text field_17" at 319,370 size 132x18; Text 'Druck-Sollw. / Pressure Setpoint'
   IOField "Template_I/O field_11" at 350,390 size 71x23; FormatPattern 99.9; Unit  Bar
      ProcessValue <- "Paramters_Paint_Mix_Pressure_Set_R"
   TextField "Template_Text field_18" at 323,270 size 125x18; Text 'Dichte-Sollw. / Density Setpoint'
   IOField "Template_I/O field_12" at 341,290 size 88x23; FormatPattern 99.9; Unit  kg/m³
      ProcessValue <- "Paramters_Paint_Mix_Density_Set_R"
   TextField "Template_Text field_19" at 475,85 size 149x23; Text 'Grünes Pigment / GREEN Pigment'
   TextField "Template_Text field_20" at 494,115 size 108x18; Text 'Füllst.-Sollw. / Level Setpoint'
   IOField "Template_I/O field_13" at 513,135 size 71x23; FormatPattern 99.9; Unit  ltr
      ProcessValue <- "Paramters_Paint_Mix_Level_Set_R"
   TextField "Template_Text field_21" at 482,166 size 133x18; Text 'Durchfluss-Sollw. / Flowrate Setpoint'
   IOField "Template_I/O field_14" at 508,186 size 80x23; FormatPattern 99.9; Unit  m³/h
      ProcessValue <- "Paramters_Paint_Mix_Flowrate_Set_R"
   TextField "Template_Text field_22" at 481,218 size 147x18; Text 'Viskositäts-Sollwert / Viscosity Setpoint'
   IOField "Template_I/O field_15" at 513,238 size 71x23; FormatPattern 99.9; Unit  cP
      ProcessValue <- "Paramters_Paint_Mix_Viscosity_Set_R"
   TextField "Template_Text field_23" at 468,320 size 161x18; Text 'Temp.-Sollwert / Temperature Setpoint'
   IOField "Template_I/O field_16" at 513,339 size 71x23; FormatPattern 99.9; Unit  °C
      ProcessValue <- "Paramters_Paint_Mix_Temperature_Set_R"
   TextField "Template_Text field_24" at 482,370 size 132x18; Text 'Druck-Sollw. / Pressure Setpoint'
   IOField "Template_I/O field_17" at 513,390 size 71x23; FormatPattern 99.9; Unit  Bar
      ProcessValue <- "Paramters_Paint_Mix_Pressure_Set_R"
   TextField "Template_Text field_25" at 486,270 size 125x18; Text 'Dichte-Sollw. / Density Setpoint'
   IOField "Template_I/O field_18" at 504,290 size 88x23; FormatPattern 99.9; Unit  kg/m³
      ProcessValue <- "Paramters_Paint_Mix_Density_Set_R"
   TextField "Template_Text field_26" at 641,85 size 146x23; Text 'Blaues Pigment / BLUE Pigment'
   TextField "Template_Text field_27" at 658,115 size 108x18; Text 'Füllst.-Sollw. / Level Setpoint'
   IOField "Template_I/O field_19" at 677,135 size 71x23; FormatPattern 99.9; Unit  ltr
      ProcessValue <- "Paramters_Paint_Mix_Level_Set_R"
   TextField "Template_Text field_28" at 646,166 size 133x18; Text 'Durchfluss-Sollw. / Flowrate Setpoint'
   IOField "Template_I/O field_20" at 672,186 size 80x23; FormatPattern 99.9; Unit  m³/h
      ProcessValue <- "Paramters_Paint_Mix_Flowrate_Set_R"
   TextField "Template_Text field_29" at 645,218 size 147x18; Text 'Viskositäts-Sollwert / Viscosity Setpoint'
   IOField "Template_I/O field_21" at 677,238 size 71x23; FormatPattern 99.9; Unit  cP
      ProcessValue <- "Paramters_Paint_Mix_Viscosity_Set_R"
   TextField "Template_Text field_30" at 632,320 size 161x18; Text 'Temp.-Sollwert / Temperature Setpoint'
   IOField "Template_I/O field_22" at 677,339 size 71x23; FormatPattern 99.9; Unit  °C
      ProcessValue <- "Paramters_Paint_Mix_Temperature_Set_R"
   TextField "Template_Text field_31" at 646,370 size 132x18; Text 'Druck-Sollw. / Pressure Setpoint'
   IOField "Template_I/O field_23" at 677,390 size 71x23; FormatPattern 99.9; Unit  Bar
      ProcessValue <- "Paramters_Paint_Mix_Pressure_Set_R"
   TextField "Template_Text field_32" at 650,270 size 125x18; Text 'Dichte-Sollw. / Density Setpoint'
   IOField "Template_I/O field_24" at 668,290 size 88x23; FormatPattern 99.9; Unit  kg/m³
      ProcessValue <- "Paramters_Paint_Mix_Density_Set_R"
   TextField "Template_Text field_33" at 78,285 size 156x23; Text 'Hauptmischb. / Main Mixer Tank'
   TextField "Template_Text field_34" at 7,319 size 166x18; Text 'Mischgeschw.-Sollw. / Mixing Speed Setpoint'
   IOField "Template_I/O field_25" at 46,339 size 88x23; FormatPattern 99.9; Unit  rpm
      ProcessValue <- "Paramters_Paint_Mix_MixingSpeed_Set_MT"
   TextField "Template_Text field_35" at 186,319 size 93x18; Text 'Aktueller pH / Current pH'
   IOField "Template_I/O field_26" at 184,339 size 88x23; FormatPattern 99.9; Unit  pH
      ProcessValue <- "Paramters_Paint_Mix_pH_MT"
   TextField "Template_Text field_36" at 23,373 size 147x18; Text 'Viskositäts-Sollwert / Viscosity Setpoint'
   IOField "Template_I/O field_27" at 46,393 size 88x23; FormatPattern 99.9; Unit  cP
      ProcessValue <- "Paramters_Paint_Mix_Viscosity_Set_MT"
   TextField "Template_Text field_37" at 174,373 size 108x18; Text 'Füllst.-Sollw. / Level Setpoint'
   IOField "Template_I/O field_28" at 184,393 size 88x23; FormatPattern 99.9; Unit  ltr
      ProcessValue <- "Paramters_Paint_Mix_Level_Set_MT"

PopupScreen "Resin_Valve_popup" 240x157
   Button "Button_1" at 27,109 size 77x35; TextOff 'ON / AN'
      on Click: SetBit("PainMix_DB_Sol_1_ValveCont"); ActivateScreen("MainOverview", 0)
      Appearance <- "PainMix_DB_Sol_1_Valve_Status"
   Button "Button_2" at 133,109 size 77x35; TextOff 'OFF / AUS'
      on Click: ResetBit("PainMix_DB_Sol_1_ValveCont"); ActivateScreen("MainOverview", 0)
      Appearance <- "PainMix_DB_Sol_1_Valve_Status"
   TextField "Text field_1" at 21,42 size 195x24; Text 'Resin Enhancer Tank / Harzverstärker-Tank'
   Button "Button_3" at 201,12 size 28x28; TextOff 'X'
      on Click: ActivateScreen("MainOverview", 0)
   TextField "Text field_2" at 44,72 size 150x23; Text 'Valve Control / Ventilsteuerung'

PopupScreen "Binder_Valve_popup" 240x157
   Button "Button_1" at 27,109 size 77x35; TextOff 'ON / AN'
      on Click: SetBit("PainMix_DB_Sol_2_ValveCont"); ActivateScreen("MainOverview", 0)
      Appearance <- "PainMix_DB_Sol_2_Valve_Status"
   Button "Button_2" at 133,109 size 77x35; TextOff 'OFF / AUS'
      on Click: ResetBit("PainMix_DB_Sol_2_ValveCont"); ActivateScreen("MainOverview", 0)
      Appearance <- "PainMix_DB_Sol_2_Valve_Status"
   Button "Button_3" at 201,12 size 28x28; TextOff 'X'
      on Click: ActivateScreen("MainOverview", 0)
   TextField "Text field_2" at 43,72 size 150x23; Text 'Valve Control / Ventilsteuerung'
   TextField "Text field_3" at 30,42 size 189x24; Text 'Solvent Binder Tank'

PopupScreen "Red_Valve_popup" 240x157
   Button "Button_1" at 27,109 size 77x35; TextOff 'ON / AN'
      on Click: SetBit("PainMix_DB_Red_ValveCont"); ActivateScreen("MainOverview", 0)
      Appearance <- "PainMix_DB_Red_Valve_Status"
   Button "Button_2" at 133,109 size 77x35; TextOff 'OFF / AUS'
      on Click: ResetBit("PainMix_DB_Red_ValveCont"); ActivateScreen("MainOverview", 0)
      Appearance <- "PainMix_DB_Red_Valve_Status"
   Button "Button_3" at 201,12 size 28x28; TextOff 'X'
      on Click: ActivateScreen("MainOverview", 0)
   TextField "Text field_2" at 44,72 size 150x23; Text 'Valve Control / Ventilsteuerung'
   TextField "Text field_1" at 26,42 size 178x24; Text 'Red Pigment Tank / Roter Pigmenttank'

PopupScreen "Green_Valve_popup" 240x157
   Button "Button_1" at 27,109 size 77x35; TextOff 'ON / AN'
      on Click: SetBit("PainMix_DB_Green_ValveCont"); ActivateScreen("MainOverview", 0)
      Appearance <- "PainMix_DB_Green_Valve_Status"
   Button "Button_2" at 133,109 size 77x35; TextOff 'OFF / AUS'
      on Click: ResetBit("PainMix_DB_Green_ValveCont"); ActivateScreen("MainOverview", 0)
      Appearance <- "PainMix_DB_Green_Valve_Status"
   Button "Button_3" at 201,12 size 28x28; TextOff 'X'
      on Click: ActivateScreen("MainOverview", 0)
   TextField "Text field_2" at 43,72 size 150x23; Text 'Valve Control / Ventilsteuerung'
   TextField "Text field_1" at 19,42 size 191x24; Text 'Green Pigment Tank / Grüner Pigmenttank'

PopupScreen "Blue_Valve_popup" 240x157
   Button "Button_1" at 27,109 size 77x35; TextOff 'ON / AN'
      on Click: SetBit("PainMix_DB_Blue_ValveCont"); ActivateScreen("MainOverview", 0)
      Appearance <- "PainMix_DB_Blue_Valve_Status"
   Button "Button_2" at 133,109 size 77x35; TextOff 'OFF / AUS'
      on Click: ResetBit("PainMix_DB_Blue_ValveCont"); ActivateScreen("MainOverview", 0)
      Appearance <- "PainMix_DB_Blue_Valve_Status"
   TextField "Text field_1" at 21,42 size 186x24; Text 'Blue Pigment Tank / Blauer Pigmenttank'
   Button "Button_3" at 201,12 size 28x28; TextOff 'X'
      on Click: ActivateScreen("MainOverview", 0)
   TextField "Text field_2" at 39,72 size 150x23; Text 'Valve Control / Ventilsteuerung'

PopupScreen "MainTank_Valve_popup" 240x157
   Button "Button_1" at 27,109 size 77x35; TextOff 'ON / AN'
      on Click: SetBit("PainMix_DB_MainTank_Mixer_Cont"); ActivateScreen("MainOverview", 0)
      Appearance <- "PainMix_DB_MainTank_Mixer_Status"
   Button "Button_2" at 133,109 size 77x35; TextOff 'OFF / AUS'
      on Click: ResetBit("PainMix_DB_MainTank_Mixer_Cont"); ActivateScreen("MainOverview", 0)
      Appearance <- "PainMix_DB_MainTank_Mixer_Status"
   TextField "Text field_1" at 38,42 size 156x24; Text 'Main Mixer Tank / Hauptmischb.'
   Button "Button_3" at 201,12 size 28x28; TextOff 'X'
      on Click: ActivateScreen("MainOverview", 0)
   TextField "Text field_2" at 43,72 size 150x23; Text 'Valve Control / Ventilsteuerung'

screen "Input_Status" 800x480, template "Inputs_temp"
   TextField "Template_Text field_2" at 300,41 size 204x25; Text 'dig. Eingänge / Digital Inputs Status'
   TextField "Text field_1" at 65,101 size 339x22; Text 'I0.0 - Resin Enhancer Level Sensor Low / I0.0 - Harzverst. Füllst.-Sens. niedrig'
   Circle "Circle_2" at 33,100 size 24x24
      Appearance <- "DI_I0.0"
   TextField "Text field_2" at 65,133 size 343x22; Text 'I0.1 - Resin Enhancer Level Sensor High / I0.1 - Harzverst. Füllst.-Sens. hoch'
   Circle "Circle_1" at 33,132 size 24x24
      Appearance <- "DI_I0.1"
   TextField "Text field_3" at 65,165 size 332x22; Text 'I0.2 - Resin Enhancer Overflow Sensor / I0.2 - Harzverst. Überlauf-Sens.'
   Circle "Circle_3" at 33,164 size 24x24
      Appearance <- "DI_I0.2"
   TextField "Text field_4" at 65,197 size 334x22; Text 'I0.3 - Solvent Binder Level Sensor Low / I0.3 - Lösb. Bind. Füllst.-Sens. niedrig'
   Circle "Circle_4" at 33,196 size 24x24
      Appearance <- "DI_I0.4"
   TextField "Text field_5" at 65,229 size 338x22; Text 'I0.4 - Solvent Binder Level Sensor High / I0.4 - Lösb. Bind. Füllst.-Sens. hoch'
   Circle "Circle_5" at 33,228 size 24x24
      Appearance <- "DI_I0.5"
   TextField "Text field_6" at 65,261 size 327x22; Text 'I0.5 - Solvent Binder Overflow Sensor / I0.5 - Lösb. Bind. Überlauf-Sens.'
   Circle "Circle_6" at 33,260 size 24x24
      Appearance <- "DI_I0.5"
   TextField "Text field_7" at 65,293 size 315x22; Text 'I0.6 - Red Pigment Level Sensor Low / I0.6 - Rotpigm. Füllst.-Sens. niedrig'
   Circle "Circle_7" at 33,292 size 24x24
      Appearance <- "DI_I0.6"
   TextField "Text field_8" at 65,325 size 319x22; Text 'I0.7 - Red Pigment Level Sensor High / I0.7 - Rotpigm. Füllst.-Sens. hoch'
   Circle "Circle_8" at 33,324 size 24x24
      Appearance <- "DI_I0.7"
   TextField "Text field_9" at 65,357 size 262x22; Text 'I1.0 - Red Pigment Valve Open / I1.0 - Rotpigm.-Vent. geöffnet'
   Circle "Circle_9" at 33,356 size 24x24
      Appearance <- "DI_I1.0"
   TextField "Text field_10" at 65,389 size 333x22; Text 'I1.1 - Green Pigment Level Sensor Low / I1.1 - Grünpigm. Füllst.-Sens. niedrig'
   Circle "Circle_10" at 33,388 size 24x24
      Appearance <- "DI_I1.1"
   Circle "Circle_11" at 428,100 size 24x24
      Appearance <- "DI_I1.2"
   TextField "Text field_12" at 460,133 size 280x22; Text 'I1.3 - Green Pigment Valve Open / I1.3 - Grünpigm.-Vent. geöffnet'
   Circle "Circle_12" at 428,132 size 24x24
      Appearance <- "DI_I1.3"
   TextField "Text field_13" at 460,165 size 320x22; Text 'I1.4 - Blue Pigment Level Sensor Low / I1.4 - Blaupigm. Füllst.-Sens. niedrig'
   Circle "Circle_13" at 428,164 size 24x24
      Appearance <- "DI_I1.4"
   TextField "Text field_14" at 460,197 size 324x22; Text 'I1.5 - Blue Pigment Level Sensor High / I1.5 - Blaupigm. Füllst.-Sens. hoch'
   Circle "Circle_14" at 428,196 size 24x24
      Appearance <- "DI_I1.5"
   TextField "Text field_15" at 460,229 size 267x22; Text 'I1.6 - Blue Pigment Valve Open / I1.6 - Blaupigm.-Vent. geöffnet'
   Circle "Circle_15" at 428,228 size 24x24
      Appearance <- "DI_I1.6"
   TextField "Text field_16" at 460,261 size 230x22; Text 'I1.7 - Agitator Running ON / I1.7 - Rührwerk läuft AN'
   Circle "Circle_16" at 428,260 size 24x24
      Appearance <- "DI_I1.7"
   TextField "Text field_17" at 460,293 size 303x22; Text 'I2.0 - Master High-Pressure Sensor / I2.0 - Haupt-Sens. Hochdruck'
   Circle "Circle_17" at 428,292 size 24x24
      Appearance <- "DI_I2.0"
   TextField "Text field_18" at 460,325 size 299x22; Text 'I2.1 - Master High-Temperature Sensor / I2.1 - Haupt-Sens. Hochtemp.'
   Circle "Circle_18" at 428,324 size 24x24
      Appearance <- "DI_I2.1"
   TextField "Text field_19" at 460,357 size 299x22; Text 'I2.2 - Master High-Temperature Sensor / I2.2 - Haupt-Sens. Hochtemp.'
   Circle "Circle_19" at 428,356 size 24x24
      Appearance <- "DI_I2.2"
   TextField "Text field_20" at 460,389 size 273x22; Text 'I2.3 - Mixing Tank Lid Open Sensor / I2.3 - Sens. Mischb. Eindeckung geöffnet'
   Circle "Circle_20" at 428,388 size 24x24
      Appearance <- "DI_I2.3"
   TextField "Text field_11" at 460,101 size 337x22; Text 'I1.2 - Green Pigment Level Sensor High / I1.2 - Grünpigm. Füllst.-Sens. hoch'

screen "Output_Status" 800x480, template "Outputs_temp"
   TextField "Template_Text field_2" at 300,41 size 207x25; Text 'dig. Ausgänge / Digital Output Status'
   TextField "Text field_1" at 65,101 size 326x22; Text 'Q0.0 - Resin Enhancer Pump Motor ON / Q0.0 - Harzverst.-Pumpenmotor AN'
   Circle "Circle_2" at 33,100 size 24x24
      Appearance <- "PainMix_DB_Sol_1_Valve_Status"
   TextField "Text field_2" at 65,133 size 337x22; Text 'Q0.1 - Resin Enhancer Inlet Valve Open / Q0.1 - Harzverst.-Einl.Vent. geöffnet'
   Circle "Circle_1" at 33,132 size 24x24
      Appearance <- "DO_Q0.1"
   TextField "Text field_3" at 65,165 size 321x22; Text 'Q0.2 - Solvent Binder Pump Motor ON / Q0.2 - Lösb. Bind.-Pumpenmotor AN'
   Circle "Circle_3" at 33,164 size 24x24
      Appearance <- "PainMix_DB_Sol_2_Valve_Status"
   TextField "Text field_4" at 65,197 size 332x22; Text 'Q0.3 - Solvent Binder Inlet Valve Open / Q0.3 - Lösb. Bind.-Einl.Vent. geöffnet'
   Circle "Circle_4" at 33,196 size 24x24
      Appearance <- "DO_Q0.3"
   TextField "Text field_5" at 65,229 size 311x22; Text 'Q0.4 - Pigment Circulation Valve ON / Q0.4 - Pigm.-Umlaufvent. AN'
   Circle "Circle_5" at 33,228 size 24x24
      Appearance <- "DO_Q0.4"
   TextField "Text field_6" at 65,261 size 302x22; Text 'Q0.5 - Red Pigment Pump Motor ON / Q0.5 - Rotpigm.-Pumpenmotor AN'
   Circle "Circle_6" at 33,260 size 24x24
      Appearance <- "PainMix_DB_Red_Valve_Status"
   TextField "Text field_7" at 65,293 size 320x22; Text 'Q0.6 - Green Pigment Pump Motor ON / Q0.6 - Grünpigm.-Pumpenmotor AN'
   Circle "Circle_7" at 33,292 size 24x24
      Appearance <- "PainMix_DB_Green_Valve_Status"
   TextField "Text field_8" at 65,325 size 307x22; Text 'Q0.7 - Blue Pigment Pump Motor ON / Q0.7 - Blaupigm.-Pumpenmotor AN'
   Circle "Circle_8" at 33,324 size 24x24
      Appearance <- "PainMix_DB_Blue_Valve_Status"
   TextField "Text field_9" at 65,357 size 276x22; Text 'Q1.0 - Pigment Inlet Valve Open / Q1.0 - Pigm.-Einl.Vent. geöffnet'
   Circle "Circle_9" at 33,356 size 24x24
      Appearance <- "DO_Q1.0"
   TextField "Text field_10" at 65,389 size 216x22; Text 'Q1.1 - Agitator Motor ON / Q1.1 - Rührw.-Motor AN'
   Circle "Circle_10" at 33,388 size 24x24
      Appearance <- "PainMix_DB_MainTank_Mixer_Status"
   Circle "Circle_11" at 428,100 size 24x24
      Appearance <- "DO_Q1.2"
   TextField "Text field_12" at 460,133 size 304x22; Text 'Q1.3 - Mixing Tank Outlet Valve ON / Q1.3 - Mischb.-Ausl.Vent. AN'
   Circle "Circle_12" at 428,132 size 24x24
      Appearance <- "DO_Q1.3"
   TextField "Text field_13" at 460,165 size 273x22; Text 'Q1.4 - Alarm Indicator Light ON / Q1.4 - Alarm-Warnl. AN'
   Circle "Circle_13" at 428,164 size 24x24
      Appearance <- "DO_Q1.4"
   TextField "Text field_14" at 460,197 size 258x22; Text 'Q1.5 - Emergency Stop Output / Q1.5 - Not-Aus-Ausg.'
   Circle "Circle_14" at 428,196 size 24x24
      Appearance <- "DO_Q1.5"
   TextField "Text field_15" at 460,229 size 255x22; Text 'Q1.6 - HMI Alarm Buzzer ON / Q1.6 - HMI-Alarm-Bummer AN'
   Circle "Circle_15" at 428,228 size 24x24
      Appearance <- "DO_Q1.6"
   TextField "Text field_16" at 460,261 size 289x22; Text 'Q1.7 - Safety Interlock Engaged ON / Q1.7 - Sicherh.-Verriegelung einger. AN'
   TextField "Text field_17" at 460,293 size 270x22; Text 'Q2.0 - Maintenance Lockout ON / Q2.0 - Wartungs-Absch. AN'
   Circle "Circle_17" at 428,292 size 24x24
      Appearance <- "DO_Q2.0"
   TextField "Text field_18" at 460,325 size 275x22; Text 'Q2.1 - Batch Complete Indicator / Q2.1 - Chargenende-Anzeige'
   Circle "Circle_18" at 428,324 size 24x24
      Appearance <- "DO_Q2.1"
   TextField "Text field_19" at 460,357 size 336x22; Text 'Q2.2 - Backup Power Actuator ON / Q2.2 - Backup-Strom-vers. Aktuator AN'
   Circle "Circle_19" at 428,356 size 24x24
      Appearance <- "DO_Q2.2"
   TextField "Text field_20" at 460,389 size 252x22; Text 'Q2.3 - Outlet Exhaust Fan ON / Q2.3 - Ausl.-Abluft-vent. AN'
   Circle "Circle_20" at 428,388 size 24x24
      Appearance <- "DO_Q2.3"
   TextField "Text field_11" at 460,101 size 297x22; Text 'Q1.2 - Mixing Tank Drain Valve ON / Q1.2 - Mischb.-Abl.Vent. AN'

Template "Outputs_temp" 800x480
   Button "Template_Button_7" at 0,1 size 799x80; TextOff 'Text'
   Button "Template_Button_6" at 560,434 size 111x44; TextOn 'Digital Inputs Dig. Eingänge'; TextOff 'Dig. Eingänge Digital Inputs'; Authorization "Monitor"
      on Click: ActivateScreen("Input_Status", 0)
      Appearance <- "Paramters_Paint_Mix_IOSt"
   GraphicView "Template_Graphic view_2" at 743,427 size 56x52; Picture "screenshot"
   Button "Template_Button_10" at 714,1 size 82x80; TextOff 'Text'
   Button "Template_Button_11" at 3,1 size 82x80; TextOff 'Text'
   GraphicView "Template_Graphic view_1" at 9,5 size 71x72; Picture "Dalle_1"
   DateTimeField "Template_Date/time field_1" at 87,37 size 107x38
   DateTimeField "Template_Date/time field_2" at 623,38 size 89x38
   Button "Template_Button_13" at 196,41 size 425x31; TextOff 'Text'
   GraphicView "Template_Graphic view_3" at 734,0 size 40x33; Picture "Graphic_4"
   Button "Template_Button_12" at 88,5 size 625x31; TextOff 'Text'
   TextField "Template_Text field_2" at 264,6 size 273x25; Text 'Farbherstellungsstation / Paint Manufacturing Station'
   Button "Button_3" at 745,424 size 53x55; TextOff 'Text'
      on Click: function_f98d16b7()
   GraphicView "Graphic view_1" at 659,5 size 53x30; Picture "Graphic_114"
      Visibility <- "Paramters_Paint_Mix_Language"
   GraphicView "Graphic view_2" at 659,5 size 53x30; Picture "Graphic_116"
      Visibility <- "Paramters_Paint_Mix_Language"
   Button "Button_7" at 650,3 size 65x37; TextOff 'Text'
      on Click: function_fb9197e8(-1)
      on Release: ResetBit("Paramters_Paint_Mix_Button_Language")
      on Press: SetBit("Paramters_Paint_Mix_Button_Language")
   IOField "Template_I/O field_1" at 717,33 size 78x24; FormatPattern ???????????????????????????????????????????????????????????????????
      ProcessValue <- "UserName_fromHMI"
   TextField "Template_Text field_1" at 716,56 size 79x21; Text 'Nutzer / Username'
   Button "Template_Button_1" at 0,434 size 111x44; TextOn 'Main Overview Hauptübersicht'; TextOff 'Hauptübersicht Main Overview'; Authorization "Monitor"
      on Click: ActivateScreen("MainOverview", 0); SetBit("Paramters_Paint_Mix_MainOverview"); ResetBit("Paramters_Paint_Mix_Parameters"); ResetBit("Paramters_Paint_Mix_RecipeM"); ResetBit("Paramters_Paint_Mix_UserM"); ResetBit("Paramters_Paint_Mix_AlarmSt"); ResetBit("Paramters_Paint_Mix_IOSt")
      Appearance <- "Paramters_Paint_Mix_MainOverview"
   Button "Template_Button_2" at 112,434 size 111x44; TextOn 'Parameter'; TextOff 'Parameter'; Authorization "Operate"
      on Click: ActivateScreen("Parameter", 0); SetBit("Paramters_Paint_Mix_Parameters"); ResetBit("Paramters_Paint_Mix_MainOverview"); ResetBit("Paramters_Paint_Mix_RecipeM"); ResetBit("Paramters_Paint_Mix_UserM"); ResetBit("Paramters_Paint_Mix_AlarmSt"); ResetBit("Paramters_Paint_Mix_IOSt")
      Appearance <- "Paramters_Paint_Mix_Parameters"
   Button "Template_Button_3" at 224,434 size 111x44; TextOn 'Recipe Management Rezept Verw.'; TextOff 'Rezept Verw. Recipe Management'; Authorization "User administration"
      on Click: ActivateScreen("Recipe", 0); SetBit("Paramters_Paint_Mix_RecipeM"); ResetBit("Paramters_Paint_Mix_Parameters"); ResetBit("Paramters_Paint_Mix_MainOverview"); ResetBit("Paramters_Paint_Mix_UserM"); ResetBit("Paramters_Paint_Mix_AlarmSt"); ResetBit("Paramters_Paint_Mix_IOSt")
      Appearance <- "Paramters_Paint_Mix_RecipeM"
   Button "Template_Button_4" at 336,434 size 111x44; TextOn 'User Management Ben. Verw.'; TextOff 'Ben. Verw. User Management'; Authorization "Monitor"
      on Click: ActivateScreen("User_Admin", 0); SetBit("Paramters_Paint_Mix_UserM"); ResetBit("Paramters_Paint_Mix_Parameters"); ResetBit("Paramters_Paint_Mix_RecipeM"); ResetBit("Paramters_Paint_Mix_MainOverview"); ResetBit("Paramters_Paint_Mix_AlarmSt"); ResetBit("Paramters_Paint_Mix_IOSt")
      Appearance <- "Paramters_Paint_Mix_UserM"
   Button "Template_Button_5" at 448,434 size 111x44; TextOn 'Alarm Status Alarm Status'; TextOff 'Alarm Status Alarm Status'; Authorization "Monitor"
      on Click: ActivateScreen("Alarm", 0); SetBit("Paramters_Paint_Mix_AlarmSt"); ResetBit("Paramters_Paint_Mix_Parameters"); ResetBit("Paramters_Paint_Mix_RecipeM"); ResetBit("Paramters_Paint_Mix_UserM"); ResetBit("Paramters_Paint_Mix_MainOverview"); ResetBit("Paramters_Paint_Mix_IOSt")
      Appearance <- "Paramters_Paint_Mix_AlarmSt"
   GraphicView "Template_Graphic view_4" at 522,411 size 43x43; Picture "Graphic_125"
      Visibility <- "Paramters_Paint_Mix_Common_A-W"

Template "Inputs_temp" 800x480
   Button "Template_Button_7" at 0,1 size 799x80; TextOff 'Text'
   Button "Template_Button_6" at 560,434 size 111x44; TextOn 'Digital Outputs Dig. Ausgänge'; TextOff 'Dig. Ausgänge Digital Outputs'; Authorization "Monitor"
      on Click: ActivateScreen("Output_Status", 0)
      Appearance <- "Paramters_Paint_Mix_IOSt"
   GraphicView "Template_Graphic view_2" at 743,427 size 56x52; Picture "screenshot"
   Button "Template_Button_10" at 714,1 size 82x80; TextOff 'Text'
   Button "Template_Button_11" at 3,1 size 82x80; TextOff 'Text'
   GraphicView "Template_Graphic view_1" at 9,5 size 71x72; Picture "Dalle_1"
   DateTimeField "Template_Date/time field_1" at 87,37 size 107x38
   DateTimeField "Template_Date/time field_2" at 623,38 size 89x38
   Button "Template_Button_13" at 196,41 size 425x31; TextOff 'Text'
   GraphicView "Template_Graphic view_3" at 734,0 size 40x33; Picture "Graphic_4"
   Button "Template_Button_12" at 88,5 size 625x31; TextOff 'Text'
   TextField "Template_Text field_2" at 264,6 size 273x25; Text 'Farbherstellungsstation / Paint Manufacturing Station'
   Button "Button_3" at 745,424 size 53x55; TextOff 'Text'
      on Click: function_f98d16b7()
   GraphicView "Graphic view_1" at 659,5 size 53x30; Picture "Graphic_114"
      Visibility <- "Paramters_Paint_Mix_Language"
   GraphicView "Graphic view_2" at 659,5 size 53x30; Picture "Graphic_116"
      Visibility <- "Paramters_Paint_Mix_Language"
   Button "Button_7" at 650,3 size 65x37; TextOff 'Text'
      on Click: function_fb9197e8(-1)
      on Release: ResetBit("Paramters_Paint_Mix_Button_Language")
      on Press: SetBit("Paramters_Paint_Mix_Button_Language")
   IOField "Template_I/O field_1" at 717,33 size 78x24; FormatPattern ???????????????????????????????????????????????????????????????????
      ProcessValue <- "UserName_fromHMI"
   TextField "Template_Text field_1" at 716,56 size 79x21; Text 'Nutzer / Username'
   Button "Template_Button_1" at 0,434 size 111x44; TextOn 'Main Overview Hauptübersicht'; TextOff 'Hauptübersicht Main Overview'; Authorization "Monitor"
      on Click: ActivateScreen("MainOverview", 0); SetBit("Paramters_Paint_Mix_MainOverview"); ResetBit("Paramters_Paint_Mix_Parameters"); ResetBit("Paramters_Paint_Mix_RecipeM"); ResetBit("Paramters_Paint_Mix_UserM"); ResetBit("Paramters_Paint_Mix_AlarmSt"); ResetBit("Paramters_Paint_Mix_IOSt")
      Appearance <- "Paramters_Paint_Mix_MainOverview"
   Button "Template_Button_2" at 112,434 size 111x44; TextOn 'Parameter'; TextOff 'Parameter'; Authorization "Operate"
      on Click: ActivateScreen("Parameter", 0); SetBit("Paramters_Paint_Mix_Parameters"); ResetBit("Paramters_Paint_Mix_MainOverview"); ResetBit("Paramters_Paint_Mix_RecipeM"); ResetBit("Paramters_Paint_Mix_UserM"); ResetBit("Paramters_Paint_Mix_AlarmSt"); ResetBit("Paramters_Paint_Mix_IOSt")
      Appearance <- "Paramters_Paint_Mix_Parameters"
   Button "Template_Button_3" at 224,434 size 111x44; TextOn 'Recipe Management Rezept Verw.'; TextOff 'Rezept Verw. Recipe Management'; Authorization "User administration"
      on Click: ActivateScreen("Recipe", 0); SetBit("Paramters_Paint_Mix_RecipeM"); ResetBit("Paramters_Paint_Mix_Parameters"); ResetBit("Paramters_Paint_Mix_MainOverview"); ResetBit("Paramters_Paint_Mix_UserM"); ResetBit("Paramters_Paint_Mix_AlarmSt"); ResetBit("Paramters_Paint_Mix_IOSt")
      Appearance <- "Paramters_Paint_Mix_RecipeM"
   Button "Template_Button_4" at 336,434 size 111x44; TextOn 'User Management Ben. Verw.'; TextOff 'Ben. Verw. User Management'; Authorization "Monitor"
      on Click: ActivateScreen("User_Admin", 0); SetBit("Paramters_Paint_Mix_UserM"); ResetBit("Paramters_Paint_Mix_Parameters"); ResetBit("Paramters_Paint_Mix_RecipeM"); ResetBit("Paramters_Paint_Mix_MainOverview"); ResetBit("Paramters_Paint_Mix_AlarmSt"); ResetBit("Paramters_Paint_Mix_IOSt")
      Appearance <- "Paramters_Paint_Mix_UserM"
   Button "Template_Button_5" at 448,434 size 111x44; TextOn 'Alarm Status Alarm Status'; TextOff 'Alarm Status Alarm Status'; Authorization "Monitor"
      on Click: ActivateScreen("Alarm", 0); SetBit("Paramters_Paint_Mix_AlarmSt"); ResetBit("Paramters_Paint_Mix_Parameters"); ResetBit("Paramters_Paint_Mix_RecipeM"); ResetBit("Paramters_Paint_Mix_UserM"); ResetBit("Paramters_Paint_Mix_MainOverview"); ResetBit("Paramters_Paint_Mix_IOSt")
      Appearance <- "Paramters_Paint_Mix_AlarmSt"
   GraphicView "Template_Graphic view_4" at 522,411 size 43x43; Picture "Graphic_125"
      Visibility <- "Paramters_Paint_Mix_Common_A-W"

screen "Recipe" 800x480, template "PaintMix"
   RecipeView "Recipe view_1" at 5,90 size 788x330; Recipe "Recipe_1"; Tag4DataRecord "Recipe_Recipe_Name"; DataRecordNameCaption 'Datensatzname: / Date Record Name:'; DataRecordNrCaption 'Nr.: / No.:'; EntryNameCaption 'Eintragsname / Entry Name'; ValueCaption 'Wert / Value'; RecipeNrCaption 'Nr.: / No.:'; RecipeNameCaption 'Rezeptname: / Recipe Name:'
   TextField "Template_Text field_2" at 315,41 size 195x25; Text 'Parameter / Recipe Management'

screen "User_Admin" 800x480, template "PaintMix"
   UserView "User view_2" at 17,90 size 754x223
   Button "Template_Button_5" at 254,353 size 118x44; TextOff 'Alarm Status / Log In'; PictureOff "Graphic_4"; PictureOn "Graphic_4"
      on Click: function_a2a04561()
   Button "Template_Button_1" at 414,353 size 118x44; TextOff 'Alarm Status / Log out'; PictureOn "Graphic_4"; PictureOff "Graphic_4"
      on Click: function_f23ef4c9()
   TextField "Template_Text field_2" at 316,41 size 175x25; Text 'dig. Eingänge / User Management'

PopupScreen "BatchDetails" 441x360
   Button "Button_1" at 110,303 size 93x35; TextOff 'MANUAL / AN'
      on Click: ResetBit("PainMix_DB_Control_Mode"); ActivateScreen("MainOverview", 0)
      Appearance <- "PainMix_DB_Control_Mode"
   Button "Button_2" at 240,303 size 93x35; TextOff 'AUTO / AUS'
      on Click: SetBit("PainMix_DB_Control_Mode"); ActivateScreen("MainOverview", 0)
      Appearance <- "PainMix_DB_Control_Mode"
   TextField "Text field_1" at 130,9 size 181x22; Text 'Recipe Details / Harzverstärker-Tank'
   Button "Button_3" at 404,8 size 28x28; TextOff 'X'
      on Click: ActivateScreen("MainOverview", 0)
   IOField "Template_I/O field_7" at 108,65 size 86x25; FormatPattern ??????????
      ProcessValue <- "Paramters_Paint_Mix_Recipe_ID"
   TextField "Text field_3" at 116,41 size 80x21; Text 'Recipe ID'
   IOField "Template_I/O field_1" at 230,65 size 105x25; FormatPattern ?????????????
      ProcessValue <- "Paramters_Paint_Mix_Recipe_Name"
   TextField "Text field_4" at 235,41 size 105x21; Text 'Recipe Name'
   TextField "Text field_2" at 130,108 size 181x22; Text 'Batch Details / Harzverstärker-Tank'
   IOField "Template_I/O field_2" at 53,164 size 86x25; FormatPattern ??????????
      ProcessValue <- "Paramters_Paint_Mix_Equip_ID"
   TextField "Text field_5" at 44,142 size 113x21; Text 'Equipment ID'
   IOField "Template_I/O field_3" at 180,164 size 86x25; FormatPattern ??????????
      ProcessValue <- "Paramters_Paint_Mix_Batch_ID"
   TextField "Text field_6" at 186,142 size 74x21; Text 'Batch ID'
   IOField "Template_I/O field_4" at 302,164 size 86x25; FormatPattern ??????????
      ProcessValue <- "Paramters_Paint_Mix_Batch_Size"
   TextField "Text field_7" at 307,142 size 86x21; Text 'Batch Size'
   IOField "Template_I/O field_5" at 124,225 size 183x25; FormatPattern ????????????????????
      ProcessValue <- "Paramters_Paint_Mix_Start_Time"
   TextField "Text field_8" at 123,203 size 185x21; Text 'Batch Start Timestamp'
   TextField "Text field_9" at 121,273 size 200x22; Text 'Control Mode Selection / Harzverstärker-Tank'

screen "Alarm" 800x480, template "PaintMix"
   TextField "Template_Text field_2" at 353,41 size 127x25; Text 'Parameter / Alarm Status'
   TextField "Template_Text field_9" at 226,95 size 211x25; Text 'Harzverstärker / Operational Warnings'
   Button "Button_8" at 662,210 size 132x44; TextOff 'Alarm Acknowledge AUS'
   Button "Button_1" at 662,278 size 132x44; TextOff 'Alarm Reset AUS'
      on Press: SetBit("PainMix_DB_Alarm_ACK")
      on Release: ResetBit("PainMix_DB_Alarm_ACK")
   TextField "Text field_7" at 6,185 size 107x38; Text 'Fill Sequence Incomplete'
   Rectangle "Rectangle_8" at 114,180 size 105x48
      Appearance <- "Paramters_Paint_Mix_Warning_2"
   TextField "Text field_8" at 117,185 size 99x38; Text 'Operator Override On'
   TextField "Text field_9" at 228,185 size 92x38; Text 'High Paint Level'
   TextField "Text field_10" at 340,185 size 82x38; Text 'Operator Inactivity'
   TextField "Text field_11" at 431,185 size 114x38; Text 'Flow Rate Inconsistency'
   TextField "Text field_12" at 551,185 size 88x38; Text 'Agitator Overspeed'
   TextField "Template_Text field_1" at 237,267 size 187x25; Text 'Harzverstärker / Operational Alarms'
   TextField "Text field_18" at 11,358 size 97x38; Text 'Filling Nozzle Leak'
   TextField "Text field_19" at 118,358 size 97x38; Text 'Emergency Stop Active'
   Rectangle "Rectangle_21" at 221,353 size 105x48
      Appearance <- "Paramters_Paint_Mix_Alarm_1"
   TextField "Text field_20" at 213,358 size 121x38; Text 'High Viscosity Detected'
   TextField "Text field_21" at 328,358 size 106x38; Text 'Mixing Tank Temperature'
   TextField "Text field_22" at 440,358 size 95x38; Text 'PLC Comm. Loss'
   TextField "Text field_23" at 539,355 size 112x38; Text 'Safety Interlock OFF'
   TextField "Text field_24" at 532,308 size 128x38; Text 'Agitator Motor Failure'
   TextField "Text field_13" at 30,308 size 60x38; Text 'Tank Overfill'
   TextField "Text field_14" at 112,308 size 110x38; Text 'Tank Overpressure'
   TextField "Text field_15" at 224,308 size 100x38; Text 'Motor Overcurrent'
   TextField "Text field_16" at 352,308 size 57x38; Text 'Valve Failure'
   Rectangle "Rectangle_17" at 435,303 size 105x48
      Appearance <- "Paramters_Paint_Mix_Alarm_2"
   TextField "Text field_17" at 450,308 size 75x38; Text 'Pump Overload'
   TextField "Text field_1" at 16,135 size 87x38; Text 'Main Tank Low Level'
   Rectangle "Rectangle_1" at 114,130 size 105x48
      Appearance <- "Paramters_Paint_Mix_Warning_1"
   TextField "Text field_2" at 113,135 size 108x38; Text 'Filter Maintenance'
   TextField "Text field_3" at 222,135 size 103x38; Text 'Agitator Maintenance'
   TextField "Text field_4" at 320,135 size 122x38; Text 'Power Backup Activated'
   TextField "Text field_5" at 439,135 size 98x38; Text 'Slow Filling Rate'
   Rectangle "Rectangle_6" at 542,130 size 105x48
      Appearance <- "Paramters_Paint_Mix_Warning_3"
   TextField "Text field_6" at 550,135 size 90x38; Text 'Nozzle Calibration'

screen "Company_Details" 800x480
   Button "Template_Button_7" at 0,1 size 799x80; TextOff 'Text'
   Button "Template_Button_11" at 3,1 size 82x80; TextOff 'Text'
   GraphicView "Template_Graphic view_1" at 9,5 size 71x72; Picture "Dalle_1"
   Button "Template_Button_12" at 88,5 size 625x31; TextOff 'Text'
   DateTimeField "Template_Date/time field_1" at 87,37 size 107x38
   Button "Template_Button_13" at 196,41 size 425x31; TextOff 'Text'
   TextField "Template_Text field_2" at 264,6 size 273x25; Text 'Farbherstellungsstation / Paint Manufacturing Station'
   TextField "Template_Text field_5" at 218,88 size 376x28; Text 'Die Welt mit Exzellenz färben / Coloring the World with Excellence'
   TextField "Template_Text field_6" at 301,41 size 215x25; Text 'Unternehmens Details / Company Details'
   GraphicView "Graphic view_1" at 425,431 size 60x38; Picture "Graphic_114"
   GraphicView "Graphic view_3" at 315,431 size 60x38; Picture "Graphic_116"
   TextField "Template_Text field_4" at 304,391 size 191x25; Text 'Sprachauswahl / Language Selection'
   Button "Button_1" at 310,425 size 69x45; TextOff 'Text'
      on Click: function_fb9197e8(-1); ResetBit("Paramters_Paint_Mix_Language")
   Button "Button_2" at 420,426 size 69x45; TextOff 'Text'
      on Click: function_fb9197e8(-1); SetBit("Paramters_Paint_Mix_Language")
   Button "Template_Button_10" at 714,1 size 82x80; TextOff 'Text'
   IOField "Template_I/O field_1" at 717,33 size 78x24; FormatPattern ????????
   GraphicView "Template_Graphic view_3" at 734,0 size 40x33; Picture "Graphic_4"
   GraphicView "Template_Graphic view_2" at 441,137 size 356x203; Picture "fuller-paint1"
   TextField "Template_Text field_3" at 2,122 size 423x211; Text 'Bei ShadeSmiths sind wir Vorreiter in innovativen Farb-Lösungen und liefern hochwertige Produkte für Industrie und Haushalt. Mit unserem Engagement für Nachhaltigkeit sorgt unsere Produktion für lebendige Farben, Haltbar Formulierungen. Entdecken Sie unser Streben nach Perfektion, und lassen jedem Untergrund Leben einhauchen. At ShadeSmiths, we are pioneers in innovative paint solutions, delivering high-quality products for industries and households. With our commitment to sustainability, our production ensures vibrant colors and durable formulations. Discover our pursuit of perfection and bring life to every surface.'
   DateTimeField "Template_Date/time field_2" at 623,38 size 89x38
   GraphicView "Graphic view_2" at 719,413 size 72x63; Picture "pngegg"
   Button "Button_3" at 720,418 size 75x55; TextOff 'Text'
      on Click: ActivateScreen("MainOverview", 0)
   TextField "Template_Text field_1" at 716,56 size 79x21; Text 'Nutzer / Username'

scheduled task "Task_1"
   on Action: function_f41c6f6c("UserName_fromHMI")
*)